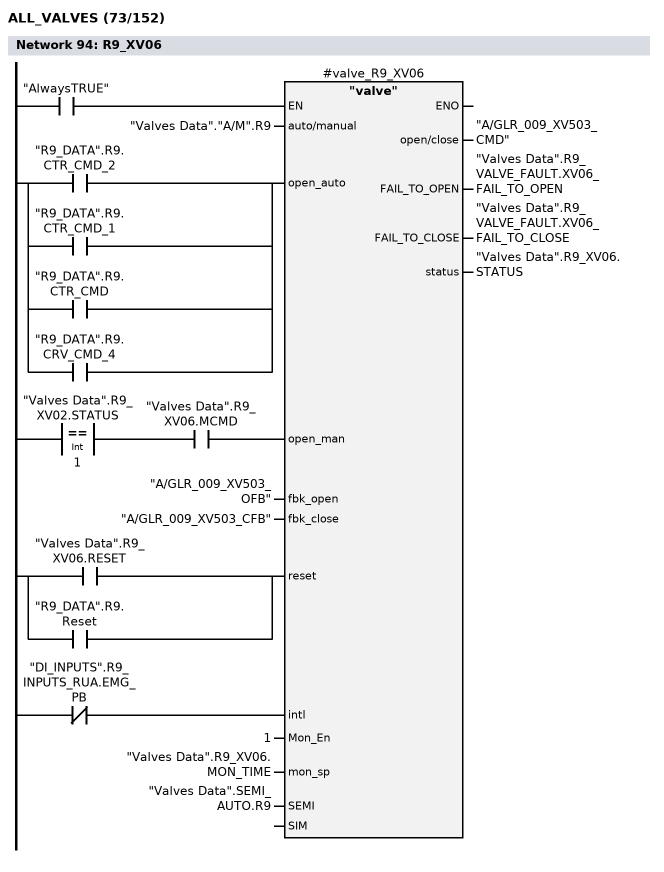
   RUNG wire#powerrail
      Contact( "AlwaysTRUE" )
      #valve_R9_XV06(open_auto := wire#w1, open_man := wire#w2, reset := wire#w3, intl := wire#w4, "auto/manual" := "Valves Data"."A/M".R9, fbk_open := "A/GLR_009_XV503_OFB", fbk_close := "A/GLR_009_XV503_CFB", Mon_En := 1, mon_sp := "Valves Data".R9_XV06.MON_TIME, SEMI := "Valves Data".SEMI_AUTO.R9, SIM :=, "open/close" => "A/GLR_009_XV503_CMD", FAIL_TO_OPEN => "Valves Data".R9_VALVE_FAULT.XV06_FAIL_TO_OPEN, FAIL_TO_CLOSE => "Valves Data".R9_VALVE_FAULT.XV06_FAIL_TO_CLOSE, status => "Valves Data".R9_XV06.STATUS)
   END_RUNG
   RUNG wire#powerrail
      Contact( "R9_DATA".R9.CTR_CMD_2 )
   END_RUNG wire#w1
   RUNG wire#powerrail
      Contact( "R9_DATA".R9.CTR_CMD_1 )
   END_RUNG wire#w1
   RUNG wire#powerrail
      Contact( "R9_DATA".R9.CTR_CMD )
   END_RUNG wire#w1
   RUNG wire#powerrail
      Contact( "R9_DATA".R9.CRV_CMD_4 )
   END_RUNG wire#w1
   RUNG wire#powerrail
      { S7_Templates := "SrcType := Int" } EQ_Contact(in1 := "Valves Data".R9_XV02.STATUS, in2 := 1)
      Contact( "Valves Data".R9_XV06.MCMD )
   END_RUNG wire#w2
   RUNG wire#powerrail
      Contact( "Valves Data".R9_XV06.RESET )
   END_RUNG wire#w3
   RUNG wire#powerrail
      Contact( "R9_DATA".R9.Reset )
   END_RUNG wire#w3
   RUNG wire#powerrail
      I_Contact( "DI_INPUTS".R9_INPUTS_RUA.EMG_PB )
   END_RUNG wire#w4
   // the same network as SCL:
   IF "AlwaysTRUE" THEN
       #valve_R9_XV06("auto/manual" := "Valves Data"."A/M".R9,   // "valve"
                      open_auto := "R9_DATA".R9.CTR_CMD_2 OR "R9_DATA".R9.CTR_CMD_1 OR "R9_DATA".R9.CTR_CMD OR "R9_DATA".R9.CRV_CMD_4,
                      open_man := ("Valves Data".R9_XV02.STATUS = 1) AND "Valves Data".R9_XV06.MCMD,
                      fbk_open := "A/GLR_009_XV503_OFB",
                      fbk_close := "A/GLR_009_XV503_CFB",
                      reset := "Valves Data".R9_XV06.RESET OR "R9_DATA".R9.Reset,
                      intl := NOT "DI_INPUTS".R9_INPUTS_RUA.EMG_PB,
                      Mon_En := 1,
                      mon_sp := "Valves Data".R9_XV06.MON_TIME,
                      SEMI := "Valves Data".SEMI_AUTO.R9,
                      "open/close" => "A/GLR_009_XV503_CMD",
                      FAIL_TO_OPEN => "Valves Data".R9_VALVE_FAULT.XV06_FAIL_TO_OPEN,
                      FAIL_TO_CLOSE => "Valves Data".R9_VALVE_FAULT.XV06_FAIL_TO_CLOSE,
                      status => "Valves Data".R9_XV06.STATUS);
   END_IF;
END_REGION

REGION Network 95: R9_XV07
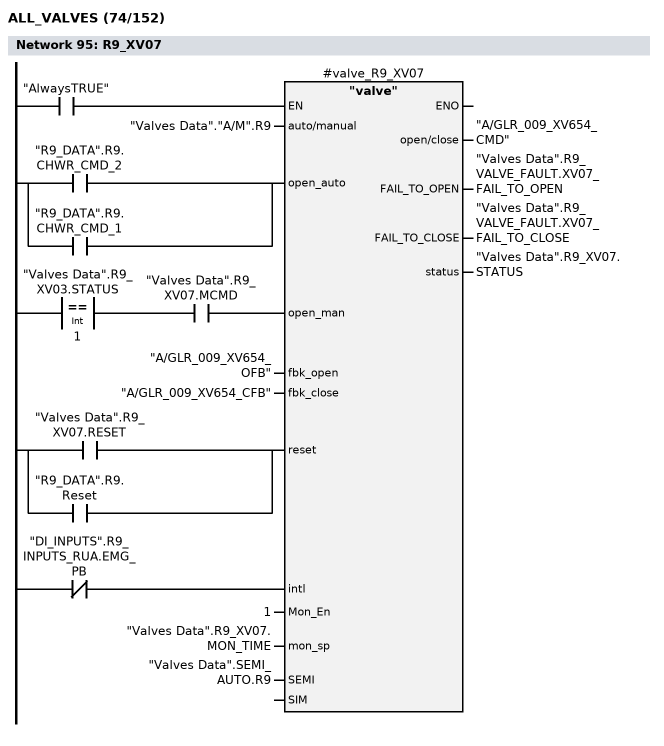
   RUNG wire#powerrail
      Contact( "AlwaysTRUE" )
      #valve_R9_XV07(open_auto := wire#w1, open_man := wire#w2, reset := wire#w3, intl := wire#w4, "auto/manual" := "Valves Data"."A/M".R9, fbk_open := "A/GLR_009_XV654_OFB", fbk_close := "A/GLR_009_XV654_CFB", Mon_En := 1, mon_sp := "Valves Data".R9_XV07.MON_TIME, SEMI := "Valves Data".SEMI_AUTO.R9, SIM :=, "open/close" => "A/GLR_009_XV654_CMD", FAIL_TO_OPEN => "Valves Data".R9_VALVE_FAULT.XV07_FAIL_TO_OPEN, FAIL_TO_CLOSE => "Valves Data".R9_VALVE_FAULT.XV07_FAIL_TO_CLOSE, status => "Valves Data".R9_XV07.STATUS)
   END_RUNG
   RUNG wire#powerrail
      Contact( "R9_DATA".R9.CHWR_CMD_2 )
   END_RUNG wire#w1
   RUNG wire#powerrail
      Contact( "R9_DATA".R9.CHWR_CMD_1 )
   END_RUNG wire#w1
   RUNG wire#powerrail
      { S7_Templates := "SrcType := Int" } EQ_Contact(in1 := "Valves Data".R9_XV03.STATUS, in2 := 1)
      Contact( "Valves Data".R9_XV07.MCMD )
   END_RUNG wire#w2
   RUNG wire#powerrail
      Contact( "Valves Data".R9_XV07.RESET )
   END_RUNG wire#w3
   RUNG wire#powerrail
      Contact( "R9_DATA".R9.Reset )
   END_RUNG wire#w3
   RUNG wire#powerrail
      I_Contact( "DI_INPUTS".R9_INPUTS_RUA.EMG_PB )
   END_RUNG wire#w4
   // the same network as SCL:
   IF "AlwaysTRUE" THEN
       #valve_R9_XV07("auto/manual" := "Valves Data"."A/M".R9,   // "valve"
                      open_auto := "R9_DATA".R9.CHWR_CMD_2 OR "R9_DATA".R9.CHWR_CMD_1,
                      open_man := ("Valves Data".R9_XV03.STATUS = 1) AND "Valves Data".R9_XV07.MCMD,
                      fbk_open := "A/GLR_009_XV654_OFB",
                      fbk_close := "A/GLR_009_XV654_CFB",
                      reset := "Valves Data".R9_XV07.RESET OR "R9_DATA".R9.Reset,
                      intl := NOT "DI_INPUTS".R9_INPUTS_RUA.EMG_PB,
                      Mon_En := 1,
                      mon_sp := "Valves Data".R9_XV07.MON_TIME,
                      SEMI := "Valves Data".SEMI_AUTO.R9,
                      "open/close" => "A/GLR_009_XV654_CMD",
                      FAIL_TO_OPEN => "Valves Data".R9_VALVE_FAULT.XV07_FAIL_TO_OPEN,
                      FAIL_TO_CLOSE => "Valves Data".R9_VALVE_FAULT.XV07_FAIL_TO_CLOSE,
                      status => "Valves Data".R9_XV07.STATUS);
   END_IF;
END_REGION

REGION Network 96: R9_XV08
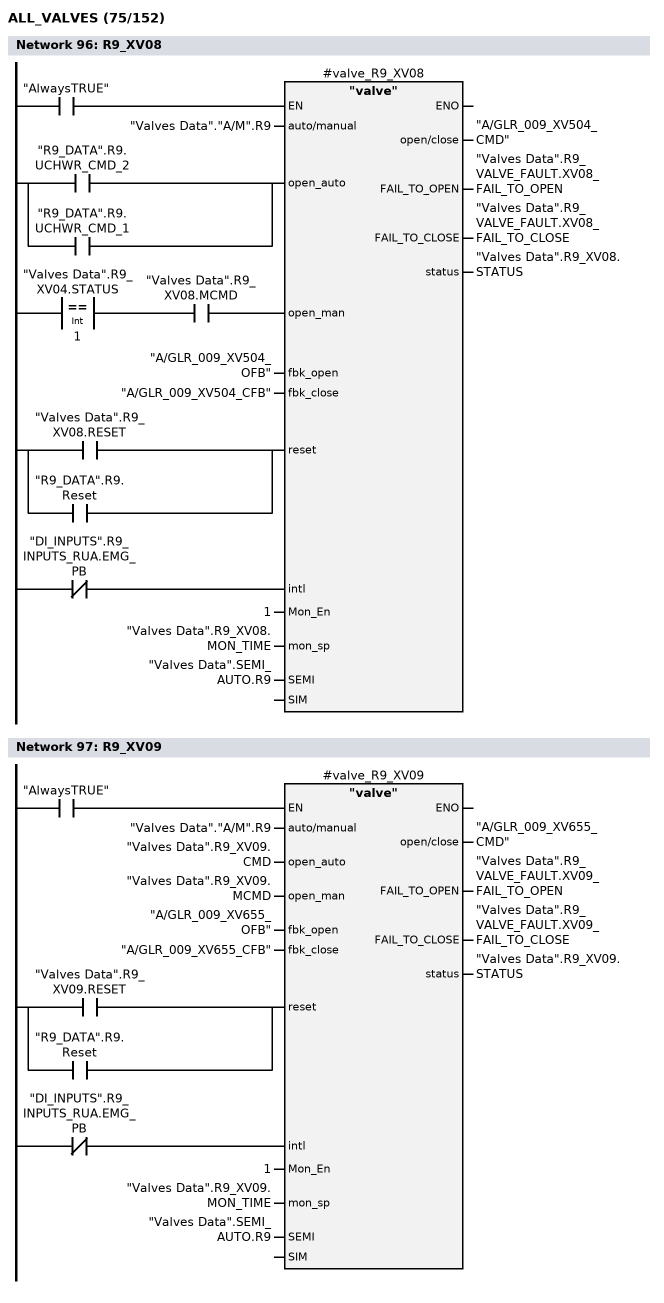
   RUNG wire#powerrail
      Contact( "AlwaysTRUE" )
      #valve_R9_XV08(open_auto := wire#w1, open_man := wire#w2, reset := wire#w3, intl := wire#w4, "auto/manual" := "Valves Data"."A/M".R9, fbk_open := "A/GLR_009_XV504_OFB", fbk_close := "A/GLR_009_XV504_CFB", Mon_En := 1, mon_sp := "Valves Data".R9_XV08.MON_TIME, SEMI := "Valves Data".SEMI_AUTO.R9, SIM :=, "open/close" => "A/GLR_009_XV504_CMD", FAIL_TO_OPEN => "Valves Data".R9_VALVE_FAULT.XV08_FAIL_TO_OPEN, FAIL_TO_CLOSE => "Valves Data".R9_VALVE_FAULT.XV08_FAIL_TO_CLOSE, status => "Valves Data".R9_XV08.STATUS)
   END_RUNG
   RUNG wire#powerrail
      Contact( "R9_DATA".R9.UCHWR_CMD_2 )
   END_RUNG wire#w1
   RUNG wire#powerrail
      Contact( "R9_DATA".R9.UCHWR_CMD_1 )
   END_RUNG wire#w1
   RUNG wire#powerrail
      { S7_Templates := "SrcType := Int" } EQ_Contact(in1 := "Valves Data".R9_XV04.STATUS, in2 := 1)
      Contact( "Valves Data".R9_XV08.MCMD )
   END_RUNG wire#w2
   RUNG wire#powerrail
      Contact( "Valves Data".R9_XV08.RESET )
   END_RUNG wire#w3
   RUNG wire#powerrail
      Contact( "R9_DATA".R9.Reset )
   END_RUNG wire#w3
   RUNG wire#powerrail
      I_Contact( "DI_INPUTS".R9_INPUTS_RUA.EMG_PB )
   END_RUNG wire#w4
   // the same network as SCL:
   IF "AlwaysTRUE" THEN
       #valve_R9_XV08("auto/manual" := "Valves Data"."A/M".R9,   // "valve"
                      open_auto := "R9_DATA".R9.UCHWR_CMD_2 OR "R9_DATA".R9.UCHWR_CMD_1,
                      open_man := ("Valves Data".R9_XV04.STATUS = 1) AND "Valves Data".R9_XV08.MCMD,
                      fbk_open := "A/GLR_009_XV504_OFB",
                      fbk_close := "A/GLR_009_XV504_CFB",
                      reset := "Valves Data".R9_XV08.RESET OR "R9_DATA".R9.Reset,
                      intl := NOT "DI_INPUTS".R9_INPUTS_RUA.EMG_PB,
                      Mon_En := 1,
                      mon_sp := "Valves Data".R9_XV08.MON_TIME,
                      SEMI := "Valves Data".SEMI_AUTO.R9,
                      "open/close" => "A/GLR_009_XV504_CMD",
                      FAIL_TO_OPEN => "Valves Data".R9_VALVE_FAULT.XV08_FAIL_TO_OPEN,
                      FAIL_TO_CLOSE => "Valves Data".R9_VALVE_FAULT.XV08_FAIL_TO_CLOSE,
                      status => "Valves Data".R9_XV08.STATUS);
   END_IF;
END_REGION

REGION Network 97: R9_XV09
   RUNG wire#powerrail
      Contact( "AlwaysTRUE" )
      #valve_R9_XV09(reset := wire#w1, intl := wire#w2, "auto/manual" := "Valves Data"."A/M".R9, open_auto := "Valves Data".R9_XV09.CMD, open_man := "Valves Data".R9_XV09.MCMD, fbk_open := "A/GLR_009_XV655_OFB", fbk_close := "A/GLR_009_XV655_CFB", Mon_En := 1, mon_sp := "Valves Data".R9_XV09.MON_TIME, SEMI := "Valves Data".SEMI_AUTO.R9, SIM :=, "open/close" => "A/GLR_009_XV655_CMD", FAIL_TO_OPEN => "Valves Data".R9_VALVE_FAULT.XV09_FAIL_TO_OPEN, FAIL_TO_CLOSE => "Valves Data".R9_VALVE_FAULT.XV09_FAIL_TO_CLOSE, status => "Valves Data".R9_XV09.STATUS)
   END_RUNG
   RUNG wire#powerrail
      Contact( "Valves Data".R9_XV09.RESET )
   END_RUNG wire#w1
   RUNG wire#powerrail
      Contact( "R9_DATA".R9.Reset )
   END_RUNG wire#w1
   RUNG wire#powerrail
      I_Contact( "DI_INPUTS".R9_INPUTS_RUA.EMG_PB )
   END_RUNG wire#w2
   // the same network as SCL:
   IF "AlwaysTRUE" THEN
       #valve_R9_XV09("auto/manual" := "Valves Data"."A/M".R9,   // "valve"
                      open_auto := "Valves Data".R9_XV09.CMD,
                      open_man := "Valves Data".R9_XV09.MCMD,
                      fbk_open := "A/GLR_009_XV655_OFB",
                      fbk_close := "A/GLR_009_XV655_CFB",
                      reset := "Valves Data".R9_XV09.RESET OR "R9_DATA".R9.Reset,
                      intl := NOT "DI_INPUTS".R9_INPUTS_RUA.EMG_PB,
                      Mon_En := 1,
                      mon_sp := "Valves Data".R9_XV09.MON_TIME,
                      SEMI := "Valves Data".SEMI_AUTO.R9,
                      "open/close" => "A/GLR_009_XV655_CMD",
                      FAIL_TO_OPEN => "Valves Data".R9_VALVE_FAULT.XV09_FAIL_TO_OPEN,
                      FAIL_TO_CLOSE => "Valves Data".R9_VALVE_FAULT.XV09_FAIL_TO_CLOSE,
                      status => "Valves Data".R9_XV09.STATUS);
   END_IF;
END_REGION

REGION Network 98: R9_XV10
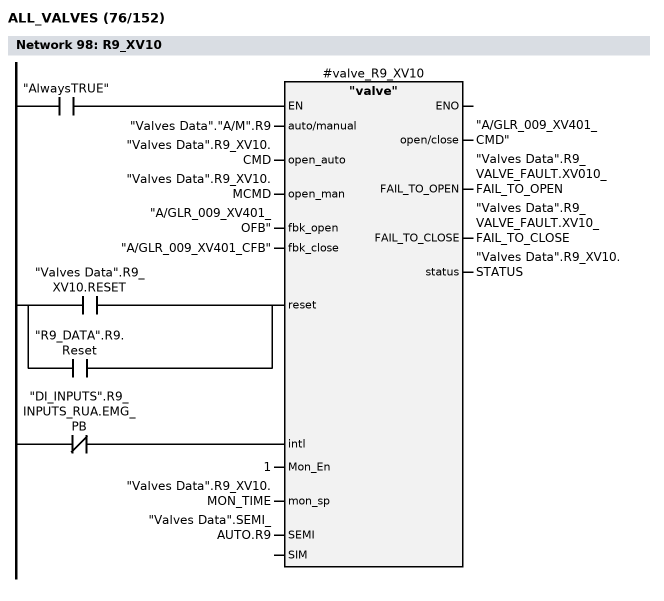
   RUNG wire#powerrail
      Contact( "AlwaysTRUE" )
      #valve_R9_XV10(reset := wire#w1, intl := wire#w2, "auto/manual" := "Valves Data"."A/M".R9, open_auto := "Valves Data".R9_XV10.CMD, open_man := "Valves Data".R9_XV10.MCMD, fbk_open := "A/GLR_009_XV401_OFB", fbk_close := "A/GLR_009_XV401_CFB", Mon_En := 1, mon_sp := "Valves Data".R9_XV10.MON_TIME, SEMI := "Valves Data".SEMI_AUTO.R9, SIM :=, "open/close" => "A/GLR_009_XV401_CMD", FAIL_TO_OPEN => "Valves Data".R9_VALVE_FAULT.XV010_FAIL_TO_OPEN, FAIL_TO_CLOSE => "Valves Data".R9_VALVE_FAULT.XV10_FAIL_TO_CLOSE, status => "Valves Data".R9_XV10.STATUS)
   END_RUNG
   RUNG wire#powerrail
      Contact( "Valves Data".R9_XV10.RESET )
   END_RUNG wire#w1
   RUNG wire#powerrail
      Contact( "R9_DATA".R9.Reset )
   END_RUNG wire#w1
   RUNG wire#powerrail
      I_Contact( "DI_INPUTS".R9_INPUTS_RUA.EMG_PB )
   END_RUNG wire#w2
   // the same network as SCL:
   IF "AlwaysTRUE" THEN
       #valve_R9_XV10("auto/manual" := "Valves Data"."A/M".R9,   // "valve"
                      open_auto := "Valves Data".R9_XV10.CMD,
                      open_man := "Valves Data".R9_XV10.MCMD,
                      fbk_open := "A/GLR_009_XV401_OFB",
                      fbk_close := "A/GLR_009_XV401_CFB",
                      reset := "Valves Data".R9_XV10.RESET OR "R9_DATA".R9.Reset,
                      intl := NOT "DI_INPUTS".R9_INPUTS_RUA.EMG_PB,
                      Mon_En := 1,
                      mon_sp := "Valves Data".R9_XV10.MON_TIME,
                      SEMI := "Valves Data".SEMI_AUTO.R9,
                      "open/close" => "A/GLR_009_XV401_CMD",
                      FAIL_TO_OPEN => "Valves Data".R9_VALVE_FAULT.XV010_FAIL_TO_OPEN,
                      FAIL_TO_CLOSE => "Valves Data".R9_VALVE_FAULT.XV10_FAIL_TO_CLOSE,
                      status => "Valves Data".R9_XV10.STATUS);
   END_IF;
END_REGION

REGION Network 99: ****REACTOR_10****
END_REGION

REGION Network 100: R10_XV01
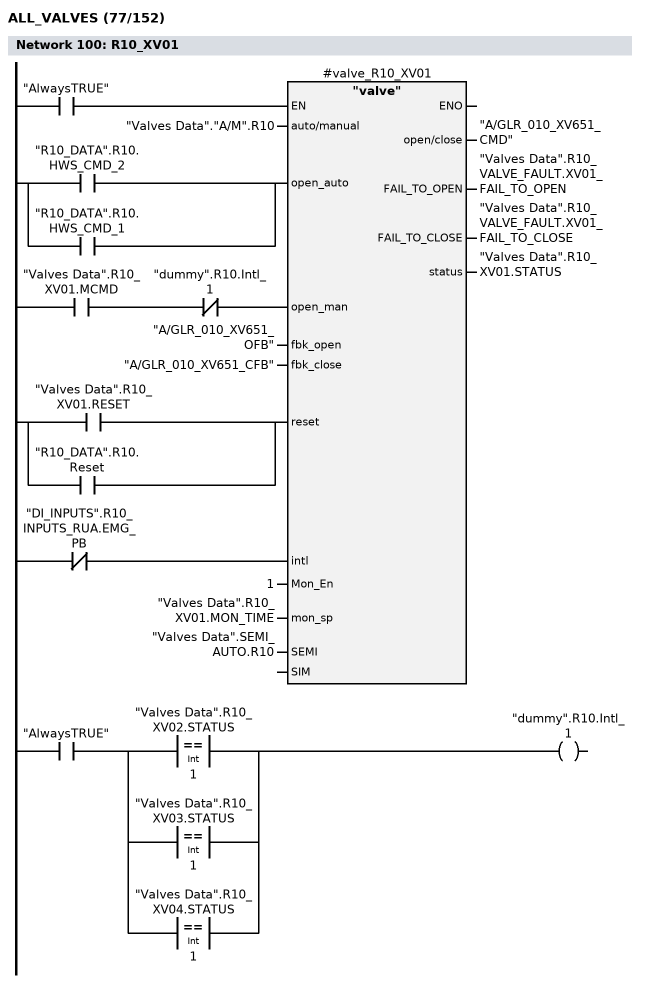
   RUNG wire#powerrail
      Contact( "AlwaysTRUE" )
      #valve_R10_XV01(open_auto := wire#w1, open_man := wire#w2, reset := wire#w3, intl := wire#w4, "auto/manual" := "Valves Data"."A/M".R10, fbk_open := "A/GLR_010_XV651_OFB", fbk_close := "A/GLR_010_XV651_CFB", Mon_En := 1, mon_sp := "Valves Data".R10_XV01.MON_TIME, SEMI := "Valves Data".SEMI_AUTO.R10, SIM :=, "open/close" => "A/GLR_010_XV651_CMD", FAIL_TO_OPEN => "Valves Data".R10_VALVE_FAULT.XV01_FAIL_TO_OPEN, FAIL_TO_CLOSE => "Valves Data".R10_VALVE_FAULT.XV01_FAIL_TO_CLOSE, status => "Valves Data".R10_XV01.STATUS)
   END_RUNG
   RUNG wire#powerrail
      Contact( "R10_DATA".R10.HWS_CMD_2 )
   END_RUNG wire#w1
   RUNG wire#powerrail
      Contact( "R10_DATA".R10.HWS_CMD_1 )
   END_RUNG wire#w1
   RUNG wire#powerrail
      Contact( "Valves Data".R10_XV01.MCMD )
      I_Contact( "dummy".R10.Intl_1 )
   END_RUNG wire#w2
   RUNG wire#powerrail
      Contact( "Valves Data".R10_XV01.RESET )
   END_RUNG wire#w3
   RUNG wire#powerrail
      Contact( "R10_DATA".R10.Reset )
   END_RUNG wire#w3
   RUNG wire#powerrail
      I_Contact( "DI_INPUTS".R10_INPUTS_RUA.EMG_PB )
   END_RUNG wire#w4
   RUNG wire#powerrail
      Contact( "AlwaysTRUE" )
      wire#w5
      { S7_Templates := "SrcType := Int" } EQ_Contact(in1 := "Valves Data".R10_XV02.STATUS, in2 := 1)
      wire#w6
      Coil( "dummy".R10.Intl_1 )
   END_RUNG
   RUNG wire#w5
      { S7_Templates := "SrcType := Int" } EQ_Contact(in1 := "Valves Data".R10_XV03.STATUS, in2 := 1)
   END_RUNG wire#w6
   RUNG wire#w5
      { S7_Templates := "SrcType := Int" } EQ_Contact(in1 := "Valves Data".R10_XV04.STATUS, in2 := 1)
   END_RUNG wire#w6
   // the same network as SCL:
   IF "AlwaysTRUE" THEN
       #valve_R10_XV01("auto/manual" := "Valves Data"."A/M".R10,   // "valve"
                       open_auto := "R10_DATA".R10.HWS_CMD_2 OR "R10_DATA".R10.HWS_CMD_1,
                       open_man := "Valves Data".R10_XV01.MCMD AND NOT "dummy".R10.Intl_1,
                       fbk_open := "A/GLR_010_XV651_OFB",
                       fbk_close := "A/GLR_010_XV651_CFB",
                       reset := "Valves Data".R10_XV01.RESET OR "R10_DATA".R10.Reset,
                       intl := NOT "DI_INPUTS".R10_INPUTS_RUA.EMG_PB,
                       Mon_En := 1,
                       mon_sp := "Valves Data".R10_XV01.MON_TIME,
                       SEMI := "Valves Data".SEMI_AUTO.R10,
                       "open/close" => "A/GLR_010_XV651_CMD",
                       FAIL_TO_OPEN => "Valves Data".R10_VALVE_FAULT.XV01_FAIL_TO_OPEN,
                       FAIL_TO_CLOSE => "Valves Data".R10_VALVE_FAULT.XV01_FAIL_TO_CLOSE,
                       status => "Valves Data".R10_XV01.STATUS);
   END_IF;
   "dummy".R10.Intl_1 := "AlwaysTRUE" AND (("Valves Data".R10_XV02.STATUS = 1) OR ("Valves Data".R10_XV03.STATUS = 1) OR ("Valves Data".R10_XV04.STATUS = 1));
END_REGION

REGION Network 101: R10_XV02
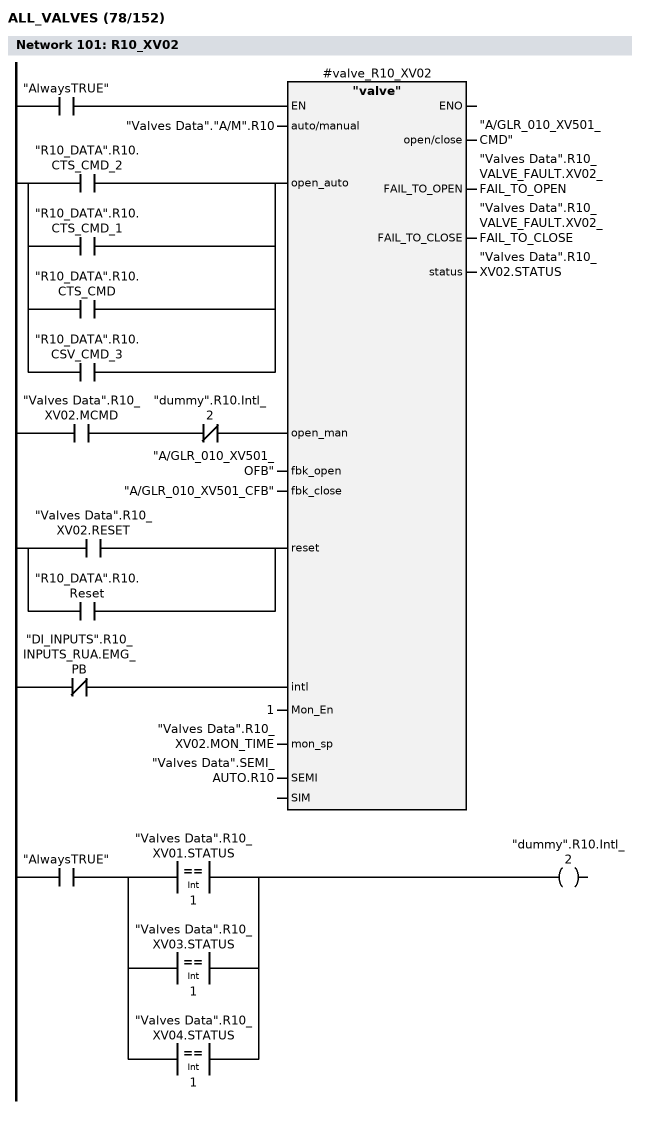
   RUNG wire#powerrail
      Contact( "AlwaysTRUE" )
      #valve_R10_XV02(open_auto := wire#w1, open_man := wire#w2, reset := wire#w3, intl := wire#w4, "auto/manual" := "Valves Data"."A/M".R10, fbk_open := "A/GLR_010_XV501_OFB", fbk_close := "A/GLR_010_XV501_CFB", Mon_En := 1, mon_sp := "Valves Data".R10_XV02.MON_TIME, SEMI := "Valves Data".SEMI_AUTO.R10, SIM :=, "open/close" => "A/GLR_010_XV501_CMD", FAIL_TO_OPEN => "Valves Data".R10_VALVE_FAULT.XV02_FAIL_TO_OPEN, FAIL_TO_CLOSE => "Valves Data".R10_VALVE_FAULT.XV02_FAIL_TO_CLOSE, status => "Valves Data".R10_XV02.STATUS)
   END_RUNG
   RUNG wire#powerrail
      Contact( "R10_DATA".R10.CTS_CMD_2 )
   END_RUNG wire#w1
   RUNG wire#powerrail
      Contact( "R10_DATA".R10.CTS_CMD_1 )
   END_RUNG wire#w1
   RUNG wire#powerrail
      Contact( "R10_DATA".R10.CTS_CMD )
   END_RUNG wire#w1
   RUNG wire#powerrail
      Contact( "R10_DATA".R10.CSV_CMD_3 )
   END_RUNG wire#w1
   RUNG wire#powerrail
      Contact( "Valves Data".R10_XV02.MCMD )
      I_Contact( "dummy".R10.Intl_2 )
   END_RUNG wire#w2
   RUNG wire#powerrail
      Contact( "Valves Data".R10_XV02.RESET )
   END_RUNG wire#w3
   RUNG wire#powerrail
      Contact( "R10_DATA".R10.Reset )
   END_RUNG wire#w3
   RUNG wire#powerrail
      I_Contact( "DI_INPUTS".R10_INPUTS_RUA.EMG_PB )
   END_RUNG wire#w4
   RUNG wire#powerrail
      Contact( "AlwaysTRUE" )
      wire#w5
      { S7_Templates := "SrcType := Int" } EQ_Contact(in1 := "Valves Data".R10_XV01.STATUS, in2 := 1)
      wire#w6
      Coil( "dummy".R10.Intl_2 )
   END_RUNG
   RUNG wire#w5
      { S7_Templates := "SrcType := Int" } EQ_Contact(in1 := "Valves Data".R10_XV03.STATUS, in2 := 1)
   END_RUNG wire#w6
   RUNG wire#w5
      { S7_Templates := "SrcType := Int" } EQ_Contact(in1 := "Valves Data".R10_XV04.STATUS, in2 := 1)
   END_RUNG wire#w6
   // the same network as SCL:
   IF "AlwaysTRUE" THEN
       #valve_R10_XV02("auto/manual" := "Valves Data"."A/M".R10,   // "valve"
                       open_auto := "R10_DATA".R10.CTS_CMD_2 OR "R10_DATA".R10.CTS_CMD_1 OR "R10_DATA".R10.CTS_CMD OR "R10_DATA".R10.CSV_CMD_3,
                       open_man := "Valves Data".R10_XV02.MCMD AND NOT "dummy".R10.Intl_2,
                       fbk_open := "A/GLR_010_XV501_OFB",
                       fbk_close := "A/GLR_010_XV501_CFB",
                       reset := "Valves Data".R10_XV02.RESET OR "R10_DATA".R10.Reset,
                       intl := NOT "DI_INPUTS".R10_INPUTS_RUA.EMG_PB,
                       Mon_En := 1,
                       mon_sp := "Valves Data".R10_XV02.MON_TIME,
                       SEMI := "Valves Data".SEMI_AUTO.R10,
                       "open/close" => "A/GLR_010_XV501_CMD",
                       FAIL_TO_OPEN => "Valves Data".R10_VALVE_FAULT.XV02_FAIL_TO_OPEN,
                       FAIL_TO_CLOSE => "Valves Data".R10_VALVE_FAULT.XV02_FAIL_TO_CLOSE,
                       status => "Valves Data".R10_XV02.STATUS);
   END_IF;
   "dummy".R10.Intl_2 := "AlwaysTRUE" AND (("Valves Data".R10_XV01.STATUS = 1) OR ("Valves Data".R10_XV03.STATUS = 1) OR ("Valves Data".R10_XV04.STATUS = 1));
END_REGION

REGION Network 102: R10_XV03
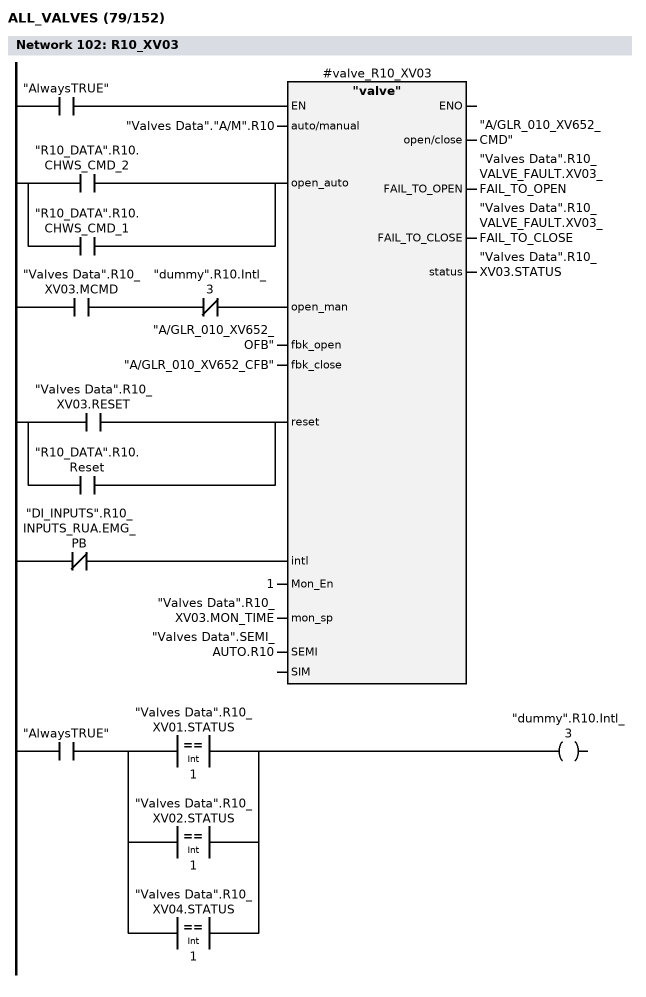
   RUNG wire#powerrail
      Contact( "AlwaysTRUE" )
      #valve_R10_XV03(open_auto := wire#w1, open_man := wire#w2, reset := wire#w3, intl := wire#w4, "auto/manual" := "Valves Data"."A/M".R10, fbk_open := "A/GLR_010_XV652_OFB", fbk_close := "A/GLR_010_XV652_CFB", Mon_En := 1, mon_sp := "Valves Data".R10_XV03.MON_TIME, SEMI := "Valves Data".SEMI_AUTO.R10, SIM :=, "open/close" => "A/GLR_010_XV652_CMD", FAIL_TO_OPEN => "Valves Data".R10_VALVE_FAULT.XV03_FAIL_TO_OPEN, FAIL_TO_CLOSE => "Valves Data".R10_VALVE_FAULT.XV03_FAIL_TO_CLOSE, status => "Valves Data".R10_XV03.STATUS)
   END_RUNG
   RUNG wire#powerrail
      Contact( "R10_DATA".R10.CHWS_CMD_2 )
   END_RUNG wire#w1
   RUNG wire#powerrail
      Contact( "R10_DATA".R10.CHWS_CMD_1 )
   END_RUNG wire#w1
   RUNG wire#powerrail
      Contact( "Valves Data".R10_XV03.MCMD )
      I_Contact( "dummy".R10.Intl_3 )
   END_RUNG wire#w2
   RUNG wire#powerrail
      Contact( "Valves Data".R10_XV03.RESET )
   END_RUNG wire#w3
   RUNG wire#powerrail
      Contact( "R10_DATA".R10.Reset )
   END_RUNG wire#w3
   RUNG wire#powerrail
      I_Contact( "DI_INPUTS".R10_INPUTS_RUA.EMG_PB )
   END_RUNG wire#w4
   RUNG wire#powerrail
      Contact( "AlwaysTRUE" )
      wire#w5
      { S7_Templates := "SrcType := Int" } EQ_Contact(in1 := "Valves Data".R10_XV01.STATUS, in2 := 1)
      wire#w6
      Coil( "dummy".R10.Intl_3 )
   END_RUNG
   RUNG wire#w5
      { S7_Templates := "SrcType := Int" } EQ_Contact(in1 := "Valves Data".R10_XV02.STATUS, in2 := 1)
   END_RUNG wire#w6
   RUNG wire#w5
      { S7_Templates := "SrcType := Int" } EQ_Contact(in1 := "Valves Data".R10_XV04.STATUS, in2 := 1)
   END_RUNG wire#w6
   // the same network as SCL:
   IF "AlwaysTRUE" THEN
       #valve_R10_XV03("auto/manual" := "Valves Data"."A/M".R10,   // "valve"
                       open_auto := "R10_DATA".R10.CHWS_CMD_2 OR "R10_DATA".R10.CHWS_CMD_1,
                       open_man := "Valves Data".R10_XV03.MCMD AND NOT "dummy".R10.Intl_3,
                       fbk_open := "A/GLR_010_XV652_OFB",
                       fbk_close := "A/GLR_010_XV652_CFB",
                       reset := "Valves Data".R10_XV03.RESET OR "R10_DATA".R10.Reset,
                       intl := NOT "DI_INPUTS".R10_INPUTS_RUA.EMG_PB,
                       Mon_En := 1,
                       mon_sp := "Valves Data".R10_XV03.MON_TIME,
                       SEMI := "Valves Data".SEMI_AUTO.R10,
                       "open/close" => "A/GLR_010_XV652_CMD",
                       FAIL_TO_OPEN => "Valves Data".R10_VALVE_FAULT.XV03_FAIL_TO_OPEN,
                       FAIL_TO_CLOSE => "Valves Data".R10_VALVE_FAULT.XV03_FAIL_TO_CLOSE,
                       status => "Valves Data".R10_XV03.STATUS);
   END_IF;
   "dummy".R10.Intl_3 := "AlwaysTRUE" AND (("Valves Data".R10_XV01.STATUS = 1) OR ("Valves Data".R10_XV02.STATUS = 1) OR ("Valves Data".R10_XV04.STATUS = 1));
END_REGION

REGION Network 103: R10_XV04
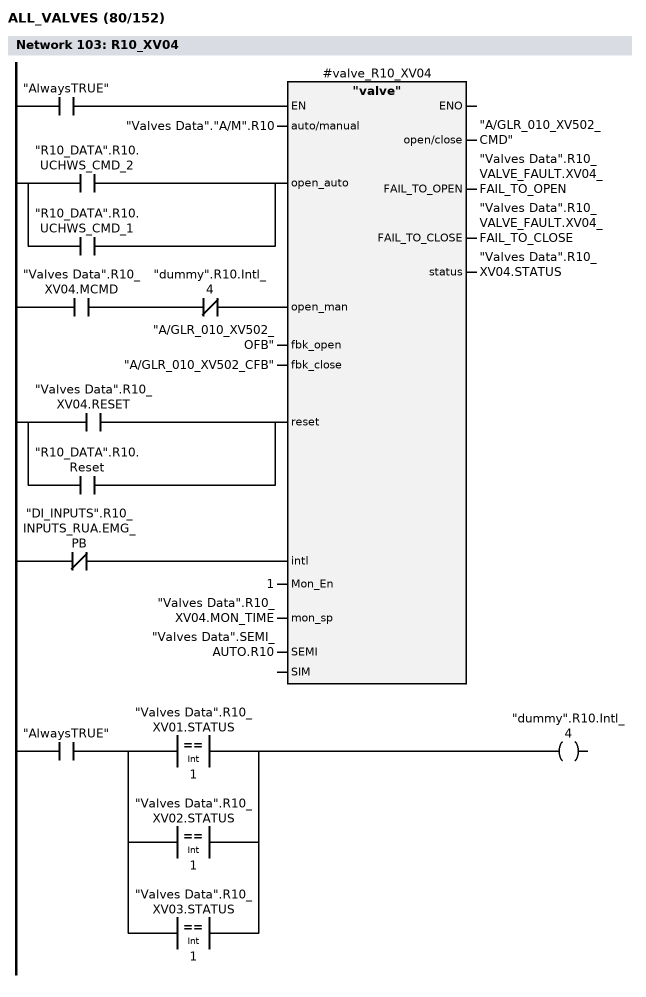
   RUNG wire#powerrail
      Contact( "AlwaysTRUE" )
      #valve_R10_XV04(open_auto := wire#w1, open_man := wire#w2, reset := wire#w3, intl := wire#w4, "auto/manual" := "Valves Data"."A/M".R10, fbk_open := "A/GLR_010_XV502_OFB", fbk_close := "A/GLR_010_XV502_CFB", Mon_En := 1, mon_sp := "Valves Data".R10_XV04.MON_TIME, SEMI := "Valves Data".SEMI_AUTO.R10, SIM :=, "open/close" => "A/GLR_010_XV502_CMD", FAIL_TO_OPEN => "Valves Data".R10_VALVE_FAULT.XV04_FAIL_TO_OPEN, FAIL_TO_CLOSE => "Valves Data".R10_VALVE_FAULT.XV04_FAIL_TO_CLOSE, status => "Valves Data".R10_XV04.STATUS)
   END_RUNG
   RUNG wire#powerrail
      Contact( "R10_DATA".R10.UCHWS_CMD_2 )
   END_RUNG wire#w1
   RUNG wire#powerrail
      Contact( "R10_DATA".R10.UCHWS_CMD_1 )
   END_RUNG wire#w1
   RUNG wire#powerrail
      Contact( "Valves Data".R10_XV04.MCMD )
      I_Contact( "dummy".R10.Intl_4 )
   END_RUNG wire#w2
   RUNG wire#powerrail
      Contact( "Valves Data".R10_XV04.RESET )
   END_RUNG wire#w3
   RUNG wire#powerrail
      Contact( "R10_DATA".R10.Reset )
   END_RUNG wire#w3
   RUNG wire#powerrail
      I_Contact( "DI_INPUTS".R10_INPUTS_RUA.EMG_PB )
   END_RUNG wire#w4
   RUNG wire#powerrail
      Contact( "AlwaysTRUE" )
      wire#w5
      { S7_Templates := "SrcType := Int" } EQ_Contact(in1 := "Valves Data".R10_XV01.STATUS, in2 := 1)
      wire#w6
      Coil( "dummy".R10.Intl_4 )
   END_RUNG
   RUNG wire#w5
      { S7_Templates := "SrcType := Int" } EQ_Contact(in1 := "Valves Data".R10_XV02.STATUS, in2 := 1)
   END_RUNG wire#w6
   RUNG wire#w5
      { S7_Templates := "SrcType := Int" } EQ_Contact(in1 := "Valves Data".R10_XV03.STATUS, in2 := 1)
   END_RUNG wire#w6
   // the same network as SCL:
   IF "AlwaysTRUE" THEN
       #valve_R10_XV04("auto/manual" := "Valves Data"."A/M".R10,   // "valve"
                       open_auto := "R10_DATA".R10.UCHWS_CMD_2 OR "R10_DATA".R10.UCHWS_CMD_1,
                       open_man := "Valves Data".R10_XV04.MCMD AND NOT "dummy".R10.Intl_4,
                       fbk_open := "A/GLR_010_XV502_OFB",
                       fbk_close := "A/GLR_010_XV502_CFB",
                       reset := "Valves Data".R10_XV04.RESET OR "R10_DATA".R10.Reset,
                       intl := NOT "DI_INPUTS".R10_INPUTS_RUA.EMG_PB,
                       Mon_En := 1,
                       mon_sp := "Valves Data".R10_XV04.MON_TIME,
                       SEMI := "Valves Data".SEMI_AUTO.R10,
                       "open/close" => "A/GLR_010_XV502_CMD",
                       FAIL_TO_OPEN => "Valves Data".R10_VALVE_FAULT.XV04_FAIL_TO_OPEN,
                       FAIL_TO_CLOSE => "Valves Data".R10_VALVE_FAULT.XV04_FAIL_TO_CLOSE,
                       status => "Valves Data".R10_XV04.STATUS);
   END_IF;
   "dummy".R10.Intl_4 := "AlwaysTRUE" AND (("Valves Data".R10_XV01.STATUS = 1) OR ("Valves Data".R10_XV02.STATUS = 1) OR ("Valves Data".R10_XV03.STATUS = 1));
END_REGION

REGION Network 104: R10_XV05
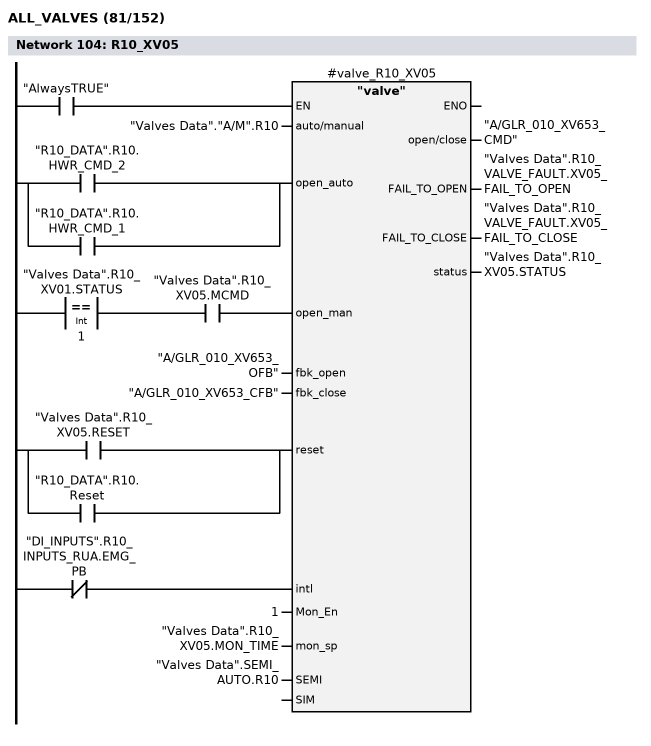
   RUNG wire#powerrail
      Contact( "AlwaysTRUE" )
      #valve_R10_XV05(open_auto := wire#w1, open_man := wire#w2, reset := wire#w3, intl := wire#w4, "auto/manual" := "Valves Data"."A/M".R10, fbk_open := "A/GLR_010_XV653_OFB", fbk_close := "A/GLR_010_XV653_CFB", Mon_En := 1, mon_sp := "Valves Data".R10_XV05.MON_TIME, SEMI := "Valves Data".SEMI_AUTO.R10, SIM :=, "open/close" => "A/GLR_010_XV653_CMD", FAIL_TO_OPEN => "Valves Data".R10_VALVE_FAULT.XV05_FAIL_TO_OPEN, FAIL_TO_CLOSE => "Valves Data".R10_VALVE_FAULT.XV05_FAIL_TO_CLOSE, status => "Valves Data".R10_XV05.STATUS)
   END_RUNG
   RUNG wire#powerrail
      Contact( "R10_DATA".R10.HWR_CMD_2 )
   END_RUNG wire#w1
   RUNG wire#powerrail
      Contact( "R10_DATA".R10.HWR_CMD_1 )
   END_RUNG wire#w1
   RUNG wire#powerrail
      { S7_Templates := "SrcType := Int" } EQ_Contact(in1 := "Valves Data".R10_XV01.STATUS, in2 := 1)
      Contact( "Valves Data".R10_XV05.MCMD )
   END_RUNG wire#w2
   RUNG wire#powerrail
      Contact( "Valves Data".R10_XV05.RESET )
   END_RUNG wire#w3
   RUNG wire#powerrail
      Contact( "R10_DATA".R10.Reset )
   END_RUNG wire#w3
   RUNG wire#powerrail
      I_Contact( "DI_INPUTS".R10_INPUTS_RUA.EMG_PB )
   END_RUNG wire#w4
   // the same network as SCL:
   IF "AlwaysTRUE" THEN
       #valve_R10_XV05("auto/manual" := "Valves Data"."A/M".R10,   // "valve"
                       open_auto := "R10_DATA".R10.HWR_CMD_2 OR "R10_DATA".R10.HWR_CMD_1,
                       open_man := ("Valves Data".R10_XV01.STATUS = 1) AND "Valves Data".R10_XV05.MCMD,
                       fbk_open := "A/GLR_010_XV653_OFB",
                       fbk_close := "A/GLR_010_XV653_CFB",
                       reset := "Valves Data".R10_XV05.RESET OR "R10_DATA".R10.Reset,
                       intl := NOT "DI_INPUTS".R10_INPUTS_RUA.EMG_PB,
                       Mon_En := 1,
                       mon_sp := "Valves Data".R10_XV05.MON_TIME,
                       SEMI := "Valves Data".SEMI_AUTO.R10,
                       "open/close" => "A/GLR_010_XV653_CMD",
                       FAIL_TO_OPEN => "Valves Data".R10_VALVE_FAULT.XV05_FAIL_TO_OPEN,
                       FAIL_TO_CLOSE => "Valves Data".R10_VALVE_FAULT.XV05_FAIL_TO_CLOSE,
                       status => "Valves Data".R10_XV05.STATUS);
   END_IF;
END_REGION

REGION Network 105: R10_XV06
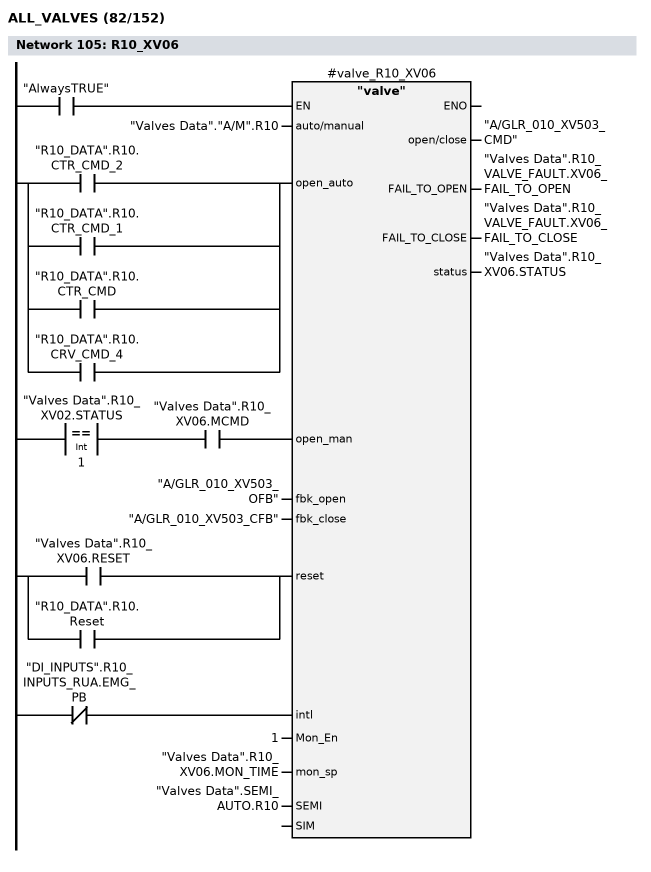
   RUNG wire#powerrail
      Contact( "AlwaysTRUE" )
      #valve_R10_XV06(open_auto := wire#w1, open_man := wire#w2, reset := wire#w3, intl := wire#w4, "auto/manual" := "Valves Data"."A/M".R10, fbk_open := "A/GLR_010_XV503_OFB", fbk_close := "A/GLR_010_XV503_CFB", Mon_En := 1, mon_sp := "Valves Data".R10_XV06.MON_TIME, SEMI := "Valves Data".SEMI_AUTO.R10, SIM :=, "open/close" => "A/GLR_010_XV503_CMD", FAIL_TO_OPEN => "Valves Data".R10_VALVE_FAULT.XV06_FAIL_TO_OPEN, FAIL_TO_CLOSE => "Valves Data".R10_VALVE_FAULT.XV06_FAIL_TO_CLOSE, status => "Valves Data".R10_XV06.STATUS)
   END_RUNG
   RUNG wire#powerrail
      Contact( "R10_DATA".R10.CTR_CMD_2 )
   END_RUNG wire#w1
   RUNG wire#powerrail
      Contact( "R10_DATA".R10.CTR_CMD_1 )
   END_RUNG wire#w1
   RUNG wire#powerrail
      Contact( "R10_DATA".R10.CTR_CMD )
   END_RUNG wire#w1
   RUNG wire#powerrail
      Contact( "R10_DATA".R10.CRV_CMD_4 )
   END_RUNG wire#w1
   RUNG wire#powerrail
      { S7_Templates := "SrcType := Int" } EQ_Contact(in1 := "Valves Data".R10_XV02.STATUS, in2 := 1)
      Contact( "Valves Data".R10_XV06.MCMD )
   END_RUNG wire#w2
   RUNG wire#powerrail
      Contact( "Valves Data".R10_XV06.RESET )
   END_RUNG wire#w3
   RUNG wire#powerrail
      Contact( "R10_DATA".R10.Reset )
   END_RUNG wire#w3
   RUNG wire#powerrail
      I_Contact( "DI_INPUTS".R10_INPUTS_RUA.EMG_PB )
   END_RUNG wire#w4
   // the same network as SCL:
   IF "AlwaysTRUE" THEN
       #valve_R10_XV06("auto/manual" := "Valves Data"."A/M".R10,   // "valve"
                       open_auto := "R10_DATA".R10.CTR_CMD_2 OR "R10_DATA".R10.CTR_CMD_1 OR "R10_DATA".R10.CTR_CMD OR "R10_DATA".R10.CRV_CMD_4,
                       open_man := ("Valves Data".R10_XV02.STATUS = 1) AND "Valves Data".R10_XV06.MCMD,
                       fbk_open := "A/GLR_010_XV503_OFB",
                       fbk_close := "A/GLR_010_XV503_CFB",
                       reset := "Valves Data".R10_XV06.RESET OR "R10_DATA".R10.Reset,
                       intl := NOT "DI_INPUTS".R10_INPUTS_RUA.EMG_PB,
                       Mon_En := 1,
                       mon_sp := "Valves Data".R10_XV06.MON_TIME,
                       SEMI := "Valves Data".SEMI_AUTO.R10,
                       "open/close" => "A/GLR_010_XV503_CMD",
                       FAIL_TO_OPEN => "Valves Data".R10_VALVE_FAULT.XV06_FAIL_TO_OPEN,
                       FAIL_TO_CLOSE => "Valves Data".R10_VALVE_FAULT.XV06_FAIL_TO_CLOSE,
                       status => "Valves Data".R10_XV06.STATUS);
   END_IF;
END_REGION

REGION Network 106: R10_XV07
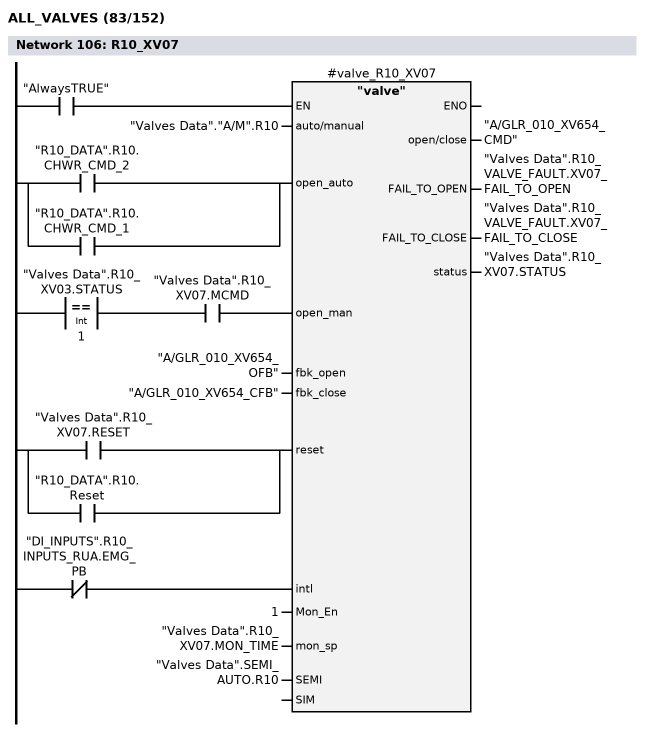
   RUNG wire#powerrail
      Contact( "AlwaysTRUE" )
      #valve_R10_XV07(open_auto := wire#w1, open_man := wire#w2, reset := wire#w3, intl := wire#w4, "auto/manual" := "Valves Data"."A/M".R10, fbk_open := "A/GLR_010_XV654_OFB", fbk_close := "A/GLR_010_XV654_CFB", Mon_En := 1, mon_sp := "Valves Data".R10_XV07.MON_TIME, SEMI := "Valves Data".SEMI_AUTO.R10, SIM :=, "open/close" => "A/GLR_010_XV654_CMD", FAIL_TO_OPEN => "Valves Data".R10_VALVE_FAULT.XV07_FAIL_TO_OPEN, FAIL_TO_CLOSE => "Valves Data".R10_VALVE_FAULT.XV07_FAIL_TO_CLOSE, status => "Valves Data".R10_XV07.STATUS)
   END_RUNG
   RUNG wire#powerrail
      Contact( "R10_DATA".R10.CHWR_CMD_2 )
   END_RUNG wire#w1
   RUNG wire#powerrail
      Contact( "R10_DATA".R10.CHWR_CMD_1 )
   END_RUNG wire#w1
   RUNG wire#powerrail
      { S7_Templates := "SrcType := Int" } EQ_Contact(in1 := "Valves Data".R10_XV03.STATUS, in2 := 1)
      Contact( "Valves Data".R10_XV07.MCMD )
   END_RUNG wire#w2
   RUNG wire#powerrail
      Contact( "Valves Data".R10_XV07.RESET )
   END_RUNG wire#w3
   RUNG wire#powerrail
      Contact( "R10_DATA".R10.Reset )
   END_RUNG wire#w3
   RUNG wire#powerrail
      I_Contact( "DI_INPUTS".R10_INPUTS_RUA.EMG_PB )
   END_RUNG wire#w4
   // the same network as SCL:
   IF "AlwaysTRUE" THEN
       #valve_R10_XV07("auto/manual" := "Valves Data"."A/M".R10,   // "valve"
                       open_auto := "R10_DATA".R10.CHWR_CMD_2 OR "R10_DATA".R10.CHWR_CMD_1,
                       open_man := ("Valves Data".R10_XV03.STATUS = 1) AND "Valves Data".R10_XV07.MCMD,
                       fbk_open := "A/GLR_010_XV654_OFB",
                       fbk_close := "A/GLR_010_XV654_CFB",
                       reset := "Valves Data".R10_XV07.RESET OR "R10_DATA".R10.Reset,
                       intl := NOT "DI_INPUTS".R10_INPUTS_RUA.EMG_PB,
                       Mon_En := 1,
                       mon_sp := "Valves Data".R10_XV07.MON_TIME,
                       SEMI := "Valves Data".SEMI_AUTO.R10,
                       "open/close" => "A/GLR_010_XV654_CMD",
                       FAIL_TO_OPEN => "Valves Data".R10_VALVE_FAULT.XV07_FAIL_TO_OPEN,
                       FAIL_TO_CLOSE => "Valves Data".R10_VALVE_FAULT.XV07_FAIL_TO_CLOSE,
                       status => "Valves Data".R10_XV07.STATUS);
   END_IF;
END_REGION

REGION Network 107: R10_XV08
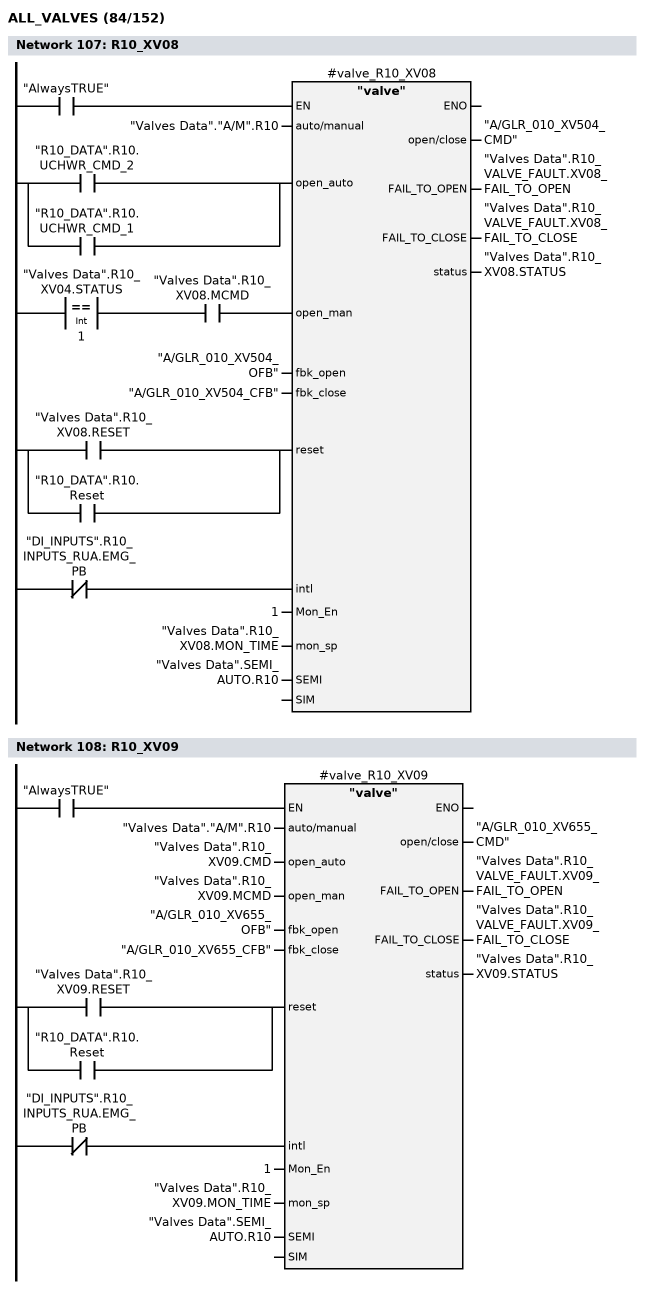
   RUNG wire#powerrail
      Contact( "AlwaysTRUE" )
      #valve_R10_XV08(open_auto := wire#w1, open_man := wire#w2, reset := wire#w3, intl := wire#w4, "auto/manual" := "Valves Data"."A/M".R10, fbk_open := "A/GLR_010_XV504_OFB", fbk_close := "A/GLR_010_XV504_CFB", Mon_En := 1, mon_sp := "Valves Data".R10_XV08.MON_TIME, SEMI := "Valves Data".SEMI_AUTO.R10, SIM :=, "open/close" => "A/GLR_010_XV504_CMD", FAIL_TO_OPEN => "Valves Data".R10_VALVE_FAULT.XV08_FAIL_TO_OPEN, FAIL_TO_CLOSE => "Valves Data".R10_VALVE_FAULT.XV08_FAIL_TO_CLOSE, status => "Valves Data".R10_XV08.STATUS)
   END_RUNG
   RUNG wire#powerrail
      Contact( "R10_DATA".R10.UCHWR_CMD_2 )
   END_RUNG wire#w1
   RUNG wire#powerrail
      Contact( "R10_DATA".R10.UCHWR_CMD_1 )
   END_RUNG wire#w1
   RUNG wire#powerrail
      { S7_Templates := "SrcType := Int" } EQ_Contact(in1 := "Valves Data".R10_XV04.STATUS, in2 := 1)
      Contact( "Valves Data".R10_XV08.MCMD )
   END_RUNG wire#w2
   RUNG wire#powerrail
      Contact( "Valves Data".R10_XV08.RESET )
   END_RUNG wire#w3
   RUNG wire#powerrail
      Contact( "R10_DATA".R10.Reset )
   END_RUNG wire#w3
   RUNG wire#powerrail
      I_Contact( "DI_INPUTS".R10_INPUTS_RUA.EMG_PB )
   END_RUNG wire#w4
   // the same network as SCL:
   IF "AlwaysTRUE" THEN
       #valve_R10_XV08("auto/manual" := "Valves Data"."A/M".R10,   // "valve"
                       open_auto := "R10_DATA".R10.UCHWR_CMD_2 OR "R10_DATA".R10.UCHWR_CMD_1,
                       open_man := ("Valves Data".R10_XV04.STATUS = 1) AND "Valves Data".R10_XV08.MCMD,
                       fbk_open := "A/GLR_010_XV504_OFB",
                       fbk_close := "A/GLR_010_XV504_CFB",
                       reset := "Valves Data".R10_XV08.RESET OR "R10_DATA".R10.Reset,
                       intl := NOT "DI_INPUTS".R10_INPUTS_RUA.EMG_PB,
                       Mon_En := 1,
                       mon_sp := "Valves Data".R10_XV08.MON_TIME,
                       SEMI := "Valves Data".SEMI_AUTO.R10,
                       "open/close" => "A/GLR_010_XV504_CMD",
                       FAIL_TO_OPEN => "Valves Data".R10_VALVE_FAULT.XV08_FAIL_TO_OPEN,
                       FAIL_TO_CLOSE => "Valves Data".R10_VALVE_FAULT.XV08_FAIL_TO_CLOSE,
                       status => "Valves Data".R10_XV08.STATUS);
   END_IF;
END_REGION

REGION Network 108: R10_XV09
   RUNG wire#powerrail
      Contact( "AlwaysTRUE" )
      #valve_R10_XV09(reset := wire#w1, intl := wire#w2, "auto/manual" := "Valves Data"."A/M".R10, open_auto := "Valves Data".R10_XV09.CMD, open_man := "Valves Data".R10_XV09.MCMD, fbk_open := "A/GLR_010_XV655_OFB", fbk_close := "A/GLR_010_XV655_CFB", Mon_En := 1, mon_sp := "Valves Data".R10_XV09.MON_TIME, SEMI := "Valves Data".SEMI_AUTO.R10, SIM :=, "open/close" => "A/GLR_010_XV655_CMD", FAIL_TO_OPEN => "Valves Data".R10_VALVE_FAULT.XV09_FAIL_TO_OPEN, FAIL_TO_CLOSE => "Valves Data".R10_VALVE_FAULT.XV09_FAIL_TO_CLOSE, status => "Valves Data".R10_XV09.STATUS)
   END_RUNG
   RUNG wire#powerrail
      Contact( "Valves Data".R10_XV09.RESET )
   END_RUNG wire#w1
   RUNG wire#powerrail
      Contact( "R10_DATA".R10.Reset )
   END_RUNG wire#w1
   RUNG wire#powerrail
      I_Contact( "DI_INPUTS".R10_INPUTS_RUA.EMG_PB )
   END_RUNG wire#w2
   // the same network as SCL:
   IF "AlwaysTRUE" THEN
       #valve_R10_XV09("auto/manual" := "Valves Data"."A/M".R10,   // "valve"
                       open_auto := "Valves Data".R10_XV09.CMD,
                       open_man := "Valves Data".R10_XV09.MCMD,
                       fbk_open := "A/GLR_010_XV655_OFB",
                       fbk_close := "A/GLR_010_XV655_CFB",
                       reset := "Valves Data".R10_XV09.RESET OR "R10_DATA".R10.Reset,
                       intl := NOT "DI_INPUTS".R10_INPUTS_RUA.EMG_PB,
                       Mon_En := 1,
                       mon_sp := "Valves Data".R10_XV09.MON_TIME,
                       SEMI := "Valves Data".SEMI_AUTO.R10,
                       "open/close" => "A/GLR_010_XV655_CMD",
                       FAIL_TO_OPEN => "Valves Data".R10_VALVE_FAULT.XV09_FAIL_TO_OPEN,
                       FAIL_TO_CLOSE => "Valves Data".R10_VALVE_FAULT.XV09_FAIL_TO_CLOSE,
                       status => "Valves Data".R10_XV09.STATUS);
   END_IF;
END_REGION

REGION Network 109: R10_XV10
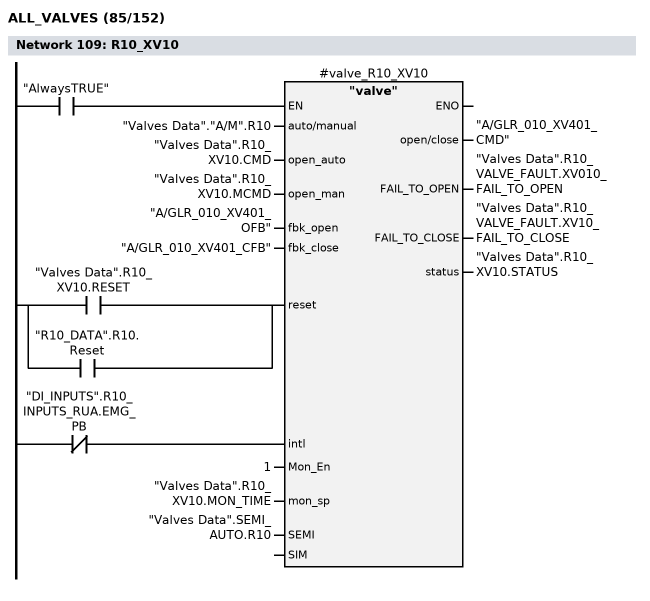
   RUNG wire#powerrail
      Contact( "AlwaysTRUE" )
      #valve_R10_XV10(reset := wire#w1, intl := wire#w2, "auto/manual" := "Valves Data"."A/M".R10, open_auto := "Valves Data".R10_XV10.CMD, open_man := "Valves Data".R10_XV10.MCMD, fbk_open := "A/GLR_010_XV401_OFB", fbk_close := "A/GLR_010_XV401_CFB", Mon_En := 1, mon_sp := "Valves Data".R10_XV10.MON_TIME, SEMI := "Valves Data".SEMI_AUTO.R10, SIM :=, "open/close" => "A/GLR_010_XV401_CMD", FAIL_TO_OPEN => "Valves Data".R10_VALVE_FAULT.XV010_FAIL_TO_OPEN, FAIL_TO_CLOSE => "Valves Data".R10_VALVE_FAULT.XV10_FAIL_TO_CLOSE, status => "Valves Data".R10_XV10.STATUS)
   END_RUNG
   RUNG wire#powerrail
      Contact( "Valves Data".R10_XV10.RESET )
   END_RUNG wire#w1
   RUNG wire#powerrail
      Contact( "R10_DATA".R10.Reset )
   END_RUNG wire#w1
   RUNG wire#powerrail
      I_Contact( "DI_INPUTS".R10_INPUTS_RUA.EMG_PB )
   END_RUNG wire#w2
   // the same network as SCL:
   IF "AlwaysTRUE" THEN
       #valve_R10_XV10("auto/manual" := "Valves Data"."A/M".R10,   // "valve"
                       open_auto := "Valves Data".R10_XV10.CMD,
                       open_man := "Valves Data".R10_XV10.MCMD,
                       fbk_open := "A/GLR_010_XV401_OFB",
                       fbk_close := "A/GLR_010_XV401_CFB",
                       reset := "Valves Data".R10_XV10.RESET OR "R10_DATA".R10.Reset,
                       intl := NOT "DI_INPUTS".R10_INPUTS_RUA.EMG_PB,
                       Mon_En := 1,
                       mon_sp := "Valves Data".R10_XV10.MON_TIME,
                       SEMI := "Valves Data".SEMI_AUTO.R10,
                       "open/close" => "A/GLR_010_XV401_CMD",
                       FAIL_TO_OPEN => "Valves Data".R10_VALVE_FAULT.XV010_FAIL_TO_OPEN,
                       FAIL_TO_CLOSE => "Valves Data".R10_VALVE_FAULT.XV10_FAIL_TO_CLOSE,
                       status => "Valves Data".R10_XV10.STATUS);
   END_IF;
END_REGION

REGION Network 110: ****REACTOR_11****
END_REGION

REGION Network 111: R11_XV01
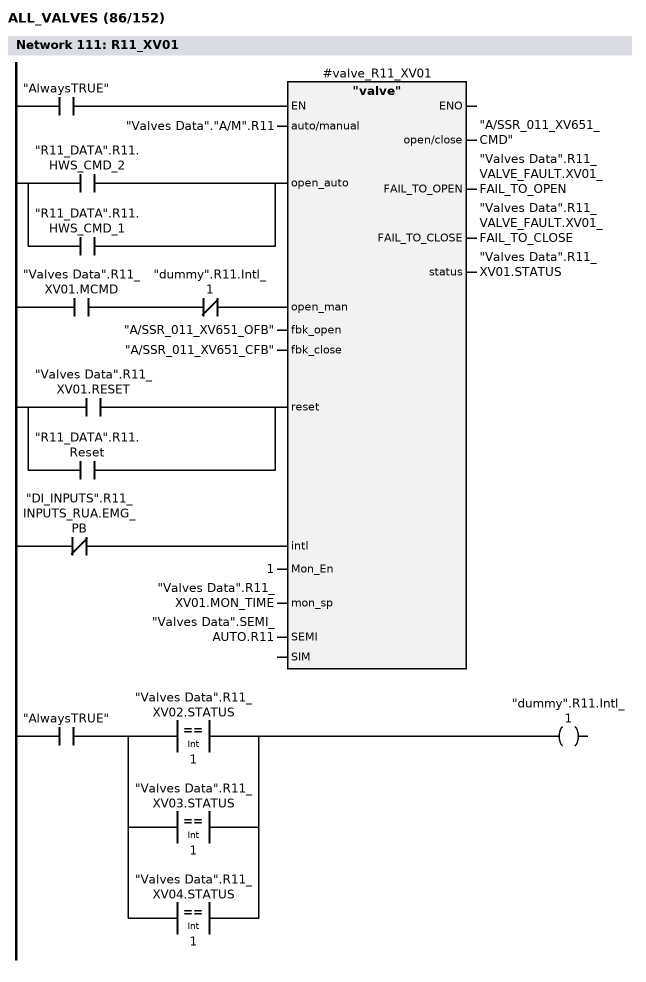
   RUNG wire#powerrail
      Contact( "AlwaysTRUE" )
      #valve_R11_XV01(open_auto := wire#w1, open_man := wire#w2, reset := wire#w3, intl := wire#w4, "auto/manual" := "Valves Data"."A/M".R11, fbk_open := "A/SSR_011_XV651_OFB", fbk_close := "A/SSR_011_XV651_CFB", Mon_En := 1, mon_sp := "Valves Data".R11_XV01.MON_TIME, SEMI := "Valves Data".SEMI_AUTO.R11, SIM :=, "open/close" => "A/SSR_011_XV651_CMD", FAIL_TO_OPEN => "Valves Data".R11_VALVE_FAULT.XV01_FAIL_TO_OPEN, FAIL_TO_CLOSE => "Valves Data".R11_VALVE_FAULT.XV01_FAIL_TO_CLOSE, status => "Valves Data".R11_XV01.STATUS)
   END_RUNG
   RUNG wire#powerrail
      Contact( "R11_DATA".R11.HWS_CMD_2 )
   END_RUNG wire#w1
   RUNG wire#powerrail
      Contact( "R11_DATA".R11.HWS_CMD_1 )
   END_RUNG wire#w1
   RUNG wire#powerrail
      Contact( "Valves Data".R11_XV01.MCMD )
      I_Contact( "dummy".R11.Intl_1 )
   END_RUNG wire#w2
   RUNG wire#powerrail
      Contact( "Valves Data".R11_XV01.RESET )
   END_RUNG wire#w3
   RUNG wire#powerrail
      Contact( "R11_DATA".R11.Reset )
   END_RUNG wire#w3
   RUNG wire#powerrail
      I_Contact( "DI_INPUTS".R11_INPUTS_RUA.EMG_PB )
   END_RUNG wire#w4
   RUNG wire#powerrail
      Contact( "AlwaysTRUE" )
      wire#w5
      { S7_Templates := "SrcType := Int" } EQ_Contact(in1 := "Valves Data".R11_XV02.STATUS, in2 := 1)
      wire#w6
      Coil( "dummy".R11.Intl_1 )
   END_RUNG
   RUNG wire#w5
      { S7_Templates := "SrcType := Int" } EQ_Contact(in1 := "Valves Data".R11_XV03.STATUS, in2 := 1)
   END_RUNG wire#w6
   RUNG wire#w5
      { S7_Templates := "SrcType := Int" } EQ_Contact(in1 := "Valves Data".R11_XV04.STATUS, in2 := 1)
   END_RUNG wire#w6
   // the same network as SCL:
   IF "AlwaysTRUE" THEN
       #valve_R11_XV01("auto/manual" := "Valves Data"."A/M".R11,   // "valve"
                       open_auto := "R11_DATA".R11.HWS_CMD_2 OR "R11_DATA".R11.HWS_CMD_1,
                       open_man := "Valves Data".R11_XV01.MCMD AND NOT "dummy".R11.Intl_1,
                       fbk_open := "A/SSR_011_XV651_OFB",
                       fbk_close := "A/SSR_011_XV651_CFB",
                       reset := "Valves Data".R11_XV01.RESET OR "R11_DATA".R11.Reset,
                       intl := NOT "DI_INPUTS".R11_INPUTS_RUA.EMG_PB,
                       Mon_En := 1,
                       mon_sp := "Valves Data".R11_XV01.MON_TIME,
                       SEMI := "Valves Data".SEMI_AUTO.R11,
                       "open/close" => "A/SSR_011_XV651_CMD",
                       FAIL_TO_OPEN => "Valves Data".R11_VALVE_FAULT.XV01_FAIL_TO_OPEN,
                       FAIL_TO_CLOSE => "Valves Data".R11_VALVE_FAULT.XV01_FAIL_TO_CLOSE,
                       status => "Valves Data".R11_XV01.STATUS);
   END_IF;
   "dummy".R11.Intl_1 := "AlwaysTRUE" AND (("Valves Data".R11_XV02.STATUS = 1) OR ("Valves Data".R11_XV03.STATUS = 1) OR ("Valves Data".R11_XV04.STATUS = 1));
END_REGION

REGION Network 112: R11_XV02
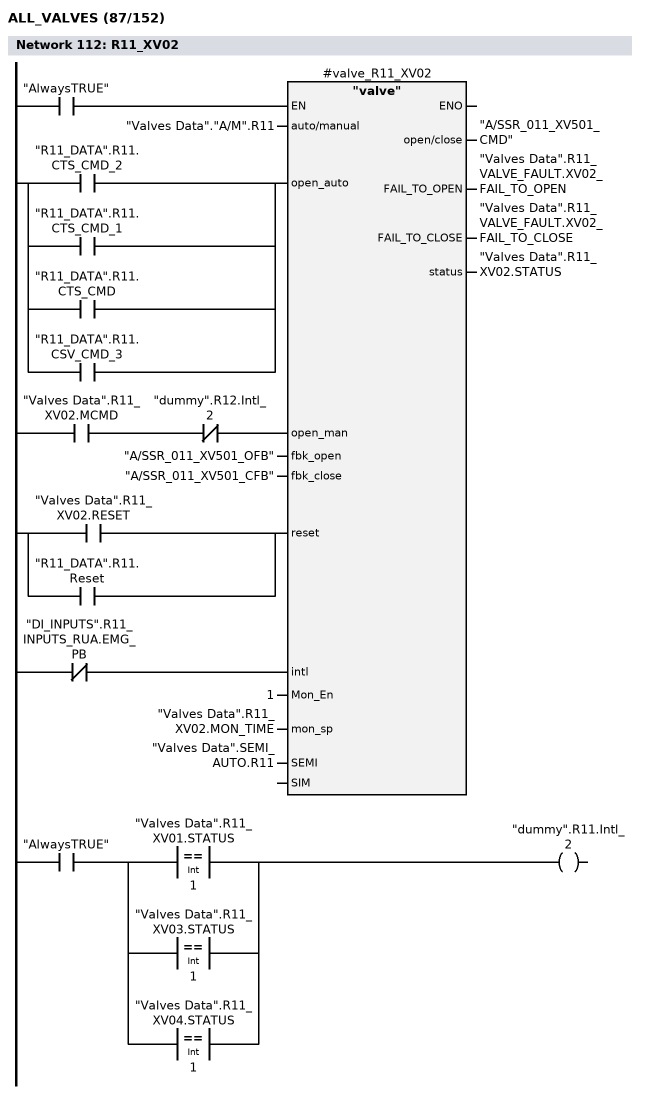
   RUNG wire#powerrail
      Contact( "AlwaysTRUE" )
      #valve_R11_XV02(open_auto := wire#w1, open_man := wire#w2, reset := wire#w3, intl := wire#w4, "auto/manual" := "Valves Data"."A/M".R11, fbk_open := "A/SSR_011_XV501_OFB", fbk_close := "A/SSR_011_XV501_CFB", Mon_En := 1, mon_sp := "Valves Data".R11_XV02.MON_TIME, SEMI := "Valves Data".SEMI_AUTO.R11, SIM :=, "open/close" => "A/SSR_011_XV501_CMD", FAIL_TO_OPEN => "Valves Data".R11_VALVE_FAULT.XV02_FAIL_TO_OPEN, FAIL_TO_CLOSE => "Valves Data".R11_VALVE_FAULT.XV02_FAIL_TO_CLOSE, status => "Valves Data".R11_XV02.STATUS)
   END_RUNG
   RUNG wire#powerrail
      Contact( "R11_DATA".R11.CTS_CMD_2 )
   END_RUNG wire#w1
   RUNG wire#powerrail
      Contact( "R11_DATA".R11.CTS_CMD_1 )
   END_RUNG wire#w1
   RUNG wire#powerrail
      Contact( "R11_DATA".R11.CTS_CMD )
   END_RUNG wire#w1
   RUNG wire#powerrail
      Contact( "R11_DATA".R11.CSV_CMD_3 )
   END_RUNG wire#w1
   RUNG wire#powerrail
      Contact( "Valves Data".R11_XV02.MCMD )
      I_Contact( "dummy".R12.Intl_2 )
   END_RUNG wire#w2
   RUNG wire#powerrail
      Contact( "Valves Data".R11_XV02.RESET )
   END_RUNG wire#w3
   RUNG wire#powerrail
      Contact( "R11_DATA".R11.Reset )
   END_RUNG wire#w3
   RUNG wire#powerrail
      I_Contact( "DI_INPUTS".R11_INPUTS_RUA.EMG_PB )
   END_RUNG wire#w4
   RUNG wire#powerrail
      Contact( "AlwaysTRUE" )
      wire#w5
      { S7_Templates := "SrcType := Int" } EQ_Contact(in1 := "Valves Data".R11_XV01.STATUS, in2 := 1)
      wire#w6
      Coil( "dummy".R11.Intl_2 )
   END_RUNG
   RUNG wire#w5
      { S7_Templates := "SrcType := Int" } EQ_Contact(in1 := "Valves Data".R11_XV03.STATUS, in2 := 1)
   END_RUNG wire#w6
   RUNG wire#w5
      { S7_Templates := "SrcType := Int" } EQ_Contact(in1 := "Valves Data".R11_XV04.STATUS, in2 := 1)
   END_RUNG wire#w6
   // the same network as SCL:
   IF "AlwaysTRUE" THEN
       #valve_R11_XV02("auto/manual" := "Valves Data"."A/M".R11,   // "valve"
                       open_auto := "R11_DATA".R11.CTS_CMD_2 OR "R11_DATA".R11.CTS_CMD_1 OR "R11_DATA".R11.CTS_CMD OR "R11_DATA".R11.CSV_CMD_3,
                       open_man := "Valves Data".R11_XV02.MCMD AND NOT "dummy".R12.Intl_2,
                       fbk_open := "A/SSR_011_XV501_OFB",
                       fbk_close := "A/SSR_011_XV501_CFB",
                       reset := "Valves Data".R11_XV02.RESET OR "R11_DATA".R11.Reset,
                       intl := NOT "DI_INPUTS".R11_INPUTS_RUA.EMG_PB,
                       Mon_En := 1,
                       mon_sp := "Valves Data".R11_XV02.MON_TIME,
                       SEMI := "Valves Data".SEMI_AUTO.R11,
                       "open/close" => "A/SSR_011_XV501_CMD",
                       FAIL_TO_OPEN => "Valves Data".R11_VALVE_FAULT.XV02_FAIL_TO_OPEN,
                       FAIL_TO_CLOSE => "Valves Data".R11_VALVE_FAULT.XV02_FAIL_TO_CLOSE,
                       status => "Valves Data".R11_XV02.STATUS);
   END_IF;
   "dummy".R11.Intl_2 := "AlwaysTRUE" AND (("Valves Data".R11_XV01.STATUS = 1) OR ("Valves Data".R11_XV03.STATUS = 1) OR ("Valves Data".R11_XV04.STATUS = 1));
END_REGION

REGION Network 113: R11_XV03
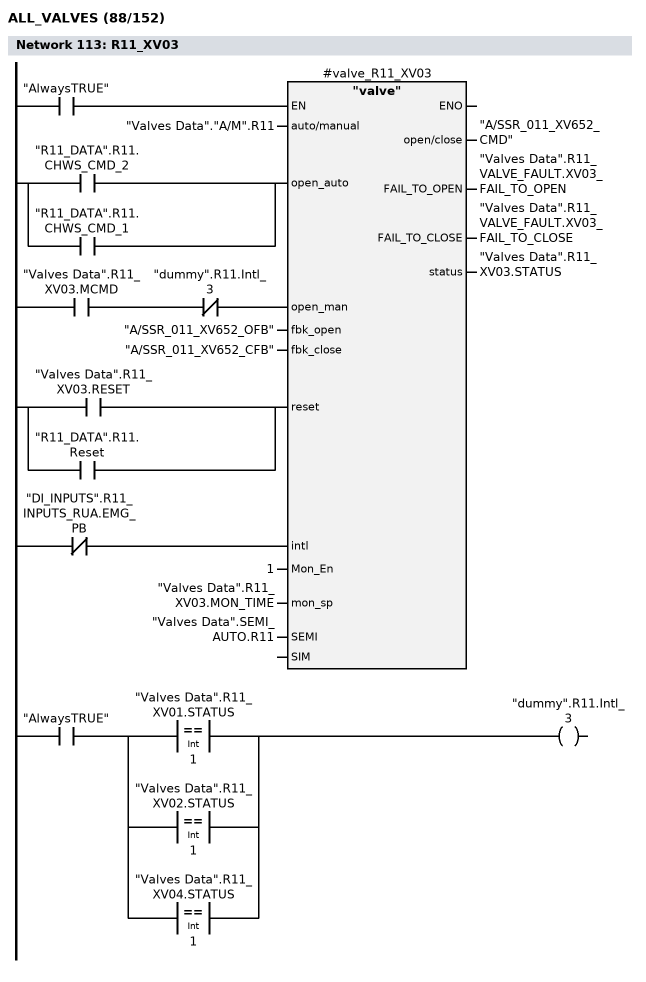
   RUNG wire#powerrail
      Contact( "AlwaysTRUE" )
      #valve_R11_XV03(open_auto := wire#w1, open_man := wire#w2, reset := wire#w3, intl := wire#w4, "auto/manual" := "Valves Data"."A/M".R11, fbk_open := "A/SSR_011_XV652_OFB", fbk_close := "A/SSR_011_XV652_CFB", Mon_En := 1, mon_sp := "Valves Data".R11_XV03.MON_TIME, SEMI := "Valves Data".SEMI_AUTO.R11, SIM :=, "open/close" => "A/SSR_011_XV652_CMD", FAIL_TO_OPEN => "Valves Data".R11_VALVE_FAULT.XV03_FAIL_TO_OPEN, FAIL_TO_CLOSE => "Valves Data".R11_VALVE_FAULT.XV03_FAIL_TO_CLOSE, status => "Valves Data".R11_XV03.STATUS)
   END_RUNG
   RUNG wire#powerrail
      Contact( "R11_DATA".R11.CHWS_CMD_2 )
   END_RUNG wire#w1
   RUNG wire#powerrail
      Contact( "R11_DATA".R11.CHWS_CMD_1 )
   END_RUNG wire#w1
   RUNG wire#powerrail
      Contact( "Valves Data".R11_XV03.MCMD )
      I_Contact( "dummy".R11.Intl_3 )
   END_RUNG wire#w2
   RUNG wire#powerrail
      Contact( "Valves Data".R11_XV03.RESET )
   END_RUNG wire#w3
   RUNG wire#powerrail
      Contact( "R11_DATA".R11.Reset )
   END_RUNG wire#w3
   RUNG wire#powerrail
      I_Contact( "DI_INPUTS".R11_INPUTS_RUA.EMG_PB )
   END_RUNG wire#w4
   RUNG wire#powerrail
      Contact( "AlwaysTRUE" )
      wire#w5
      { S7_Templates := "SrcType := Int" } EQ_Contact(in1 := "Valves Data".R11_XV01.STATUS, in2 := 1)
      wire#w6
      Coil( "dummy".R11.Intl_3 )
   END_RUNG
   RUNG wire#w5
      { S7_Templates := "SrcType := Int" } EQ_Contact(in1 := "Valves Data".R11_XV02.STATUS, in2 := 1)
   END_RUNG wire#w6
   RUNG wire#w5
      { S7_Templates := "SrcType := Int" } EQ_Contact(in1 := "Valves Data".R11_XV04.STATUS, in2 := 1)
   END_RUNG wire#w6
   // the same network as SCL:
   IF "AlwaysTRUE" THEN
       #valve_R11_XV03("auto/manual" := "Valves Data"."A/M".R11,   // "valve"
                       open_auto := "R11_DATA".R11.CHWS_CMD_2 OR "R11_DATA".R11.CHWS_CMD_1,
                       open_man := "Valves Data".R11_XV03.MCMD AND NOT "dummy".R11.Intl_3,
                       fbk_open := "A/SSR_011_XV652_OFB",
                       fbk_close := "A/SSR_011_XV652_CFB",
                       reset := "Valves Data".R11_XV03.RESET OR "R11_DATA".R11.Reset,
                       intl := NOT "DI_INPUTS".R11_INPUTS_RUA.EMG_PB,
                       Mon_En := 1,
                       mon_sp := "Valves Data".R11_XV03.MON_TIME,
                       SEMI := "Valves Data".SEMI_AUTO.R11,
                       "open/close" => "A/SSR_011_XV652_CMD",
                       FAIL_TO_OPEN => "Valves Data".R11_VALVE_FAULT.XV03_FAIL_TO_OPEN,
                       FAIL_TO_CLOSE => "Valves Data".R11_VALVE_FAULT.XV03_FAIL_TO_CLOSE,
                       status => "Valves Data".R11_XV03.STATUS);
   END_IF;
   "dummy".R11.Intl_3 := "AlwaysTRUE" AND (("Valves Data".R11_XV01.STATUS = 1) OR ("Valves Data".R11_XV02.STATUS = 1) OR ("Valves Data".R11_XV04.STATUS = 1));
END_REGION

REGION Network 114: R11_XV04
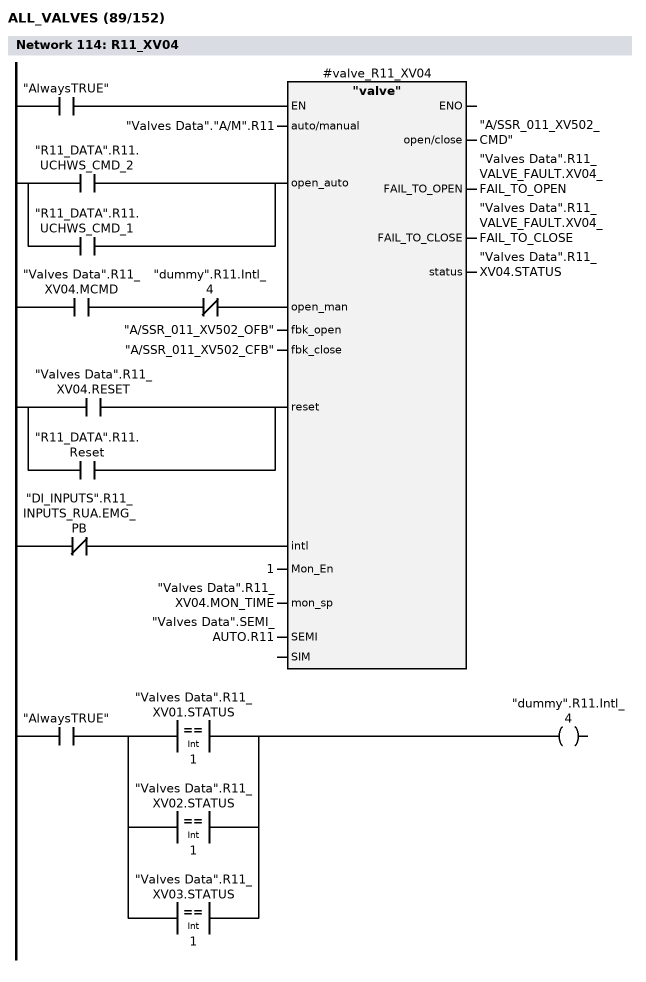
   RUNG wire#powerrail
      Contact( "AlwaysTRUE" )
      #valve_R11_XV04(open_auto := wire#w1, open_man := wire#w2, reset := wire#w3, intl := wire#w4, "auto/manual" := "Valves Data"."A/M".R11, fbk_open := "A/SSR_011_XV502_OFB", fbk_close := "A/SSR_011_XV502_CFB", Mon_En := 1, mon_sp := "Valves Data".R11_XV04.MON_TIME, SEMI := "Valves Data".SEMI_AUTO.R11, SIM :=, "open/close" => "A/SSR_011_XV502_CMD", FAIL_TO_OPEN => "Valves Data".R11_VALVE_FAULT.XV04_FAIL_TO_OPEN, FAIL_TO_CLOSE => "Valves Data".R11_VALVE_FAULT.XV04_FAIL_TO_CLOSE, status => "Valves Data".R11_XV04.STATUS)
   END_RUNG
   RUNG wire#powerrail
      Contact( "R11_DATA".R11.UCHWS_CMD_2 )
   END_RUNG wire#w1
   RUNG wire#powerrail
      Contact( "R11_DATA".R11.UCHWS_CMD_1 )
   END_RUNG wire#w1
   RUNG wire#powerrail
      Contact( "Valves Data".R11_XV04.MCMD )
      I_Contact( "dummy".R11.Intl_4 )
   END_RUNG wire#w2
   RUNG wire#powerrail
      Contact( "Valves Data".R11_XV04.RESET )
   END_RUNG wire#w3
   RUNG wire#powerrail
      Contact( "R11_DATA".R11.Reset )
   END_RUNG wire#w3
   RUNG wire#powerrail
      I_Contact( "DI_INPUTS".R11_INPUTS_RUA.EMG_PB )
   END_RUNG wire#w4
   RUNG wire#powerrail
      Contact( "AlwaysTRUE" )
      wire#w5
      { S7_Templates := "SrcType := Int" } EQ_Contact(in1 := "Valves Data".R11_XV01.STATUS, in2 := 1)
      wire#w6
      Coil( "dummy".R11.Intl_4 )
   END_RUNG
   RUNG wire#w5
      { S7_Templates := "SrcType := Int" } EQ_Contact(in1 := "Valves Data".R11_XV02.STATUS, in2 := 1)
   END_RUNG wire#w6
   RUNG wire#w5
      { S7_Templates := "SrcType := Int" } EQ_Contact(in1 := "Valves Data".R11_XV03.STATUS, in2 := 1)
   END_RUNG wire#w6
   // the same network as SCL:
   IF "AlwaysTRUE" THEN
       #valve_R11_XV04("auto/manual" := "Valves Data"."A/M".R11,   // "valve"
                       open_auto := "R11_DATA".R11.UCHWS_CMD_2 OR "R11_DATA".R11.UCHWS_CMD_1,
                       open_man := "Valves Data".R11_XV04.MCMD AND NOT "dummy".R11.Intl_4,
                       fbk_open := "A/SSR_011_XV502_OFB",
                       fbk_close := "A/SSR_011_XV502_CFB",
                       reset := "Valves Data".R11_XV04.RESET OR "R11_DATA".R11.Reset,
                       intl := NOT "DI_INPUTS".R11_INPUTS_RUA.EMG_PB,
                       Mon_En := 1,
                       mon_sp := "Valves Data".R11_XV04.MON_TIME,
                       SEMI := "Valves Data".SEMI_AUTO.R11,
                       "open/close" => "A/SSR_011_XV502_CMD",
                       FAIL_TO_OPEN => "Valves Data".R11_VALVE_FAULT.XV04_FAIL_TO_OPEN,
                       FAIL_TO_CLOSE => "Valves Data".R11_VALVE_FAULT.XV04_FAIL_TO_CLOSE,
                       status => "Valves Data".R11_XV04.STATUS);
   END_IF;
   "dummy".R11.Intl_4 := "AlwaysTRUE" AND (("Valves Data".R11_XV01.STATUS = 1) OR ("Valves Data".R11_XV02.STATUS = 1) OR ("Valves Data".R11_XV03.STATUS = 1));
END_REGION

REGION Network 115: R11_XV05
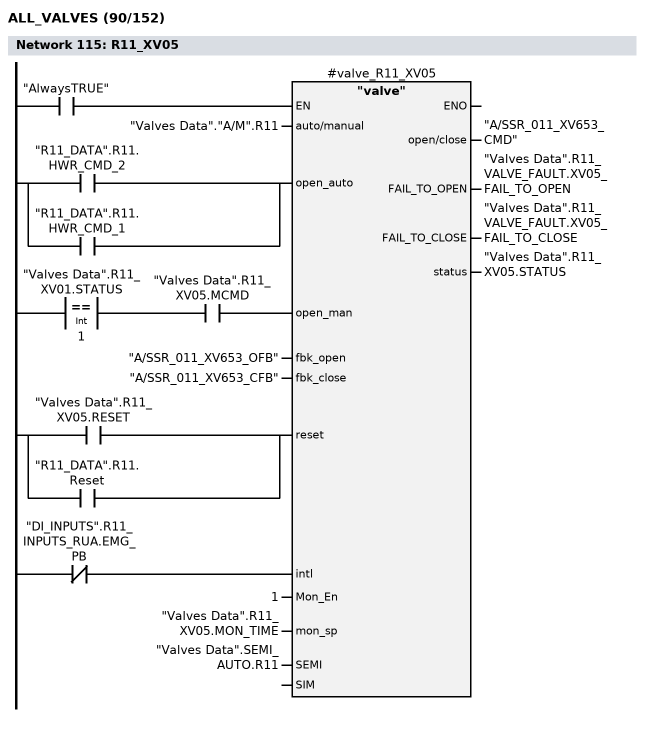
   RUNG wire#powerrail
      Contact( "AlwaysTRUE" )
      #valve_R11_XV05(open_auto := wire#w1, open_man := wire#w2, reset := wire#w3, intl := wire#w4, "auto/manual" := "Valves Data"."A/M".R11, fbk_open := "A/SSR_011_XV653_OFB", fbk_close := "A/SSR_011_XV653_CFB", Mon_En := 1, mon_sp := "Valves Data".R11_XV05.MON_TIME, SEMI := "Valves Data".SEMI_AUTO.R11, SIM :=, "open/close" => "A/SSR_011_XV653_CMD", FAIL_TO_OPEN => "Valves Data".R11_VALVE_FAULT.XV05_FAIL_TO_OPEN, FAIL_TO_CLOSE => "Valves Data".R11_VALVE_FAULT.XV05_FAIL_TO_CLOSE, status => "Valves Data".R11_XV05.STATUS)
   END_RUNG
   RUNG wire#powerrail
      Contact( "R11_DATA".R11.HWR_CMD_2 )
   END_RUNG wire#w1
   RUNG wire#powerrail
      Contact( "R11_DATA".R11.HWR_CMD_1 )
   END_RUNG wire#w1
   RUNG wire#powerrail
      { S7_Templates := "SrcType := Int" } EQ_Contact(in1 := "Valves Data".R11_XV01.STATUS, in2 := 1)
      Contact( "Valves Data".R11_XV05.MCMD )
   END_RUNG wire#w2
   RUNG wire#powerrail
      Contact( "Valves Data".R11_XV05.RESET )
   END_RUNG wire#w3
   RUNG wire#powerrail
      Contact( "R11_DATA".R11.Reset )
   END_RUNG wire#w3
   RUNG wire#powerrail
      I_Contact( "DI_INPUTS".R11_INPUTS_RUA.EMG_PB )
   END_RUNG wire#w4
   // the same network as SCL:
   IF "AlwaysTRUE" THEN
       #valve_R11_XV05("auto/manual" := "Valves Data"."A/M".R11,   // "valve"
                       open_auto := "R11_DATA".R11.HWR_CMD_2 OR "R11_DATA".R11.HWR_CMD_1,
                       open_man := ("Valves Data".R11_XV01.STATUS = 1) AND "Valves Data".R11_XV05.MCMD,
                       fbk_open := "A/SSR_011_XV653_OFB",
                       fbk_close := "A/SSR_011_XV653_CFB",
                       reset := "Valves Data".R11_XV05.RESET OR "R11_DATA".R11.Reset,
                       intl := NOT "DI_INPUTS".R11_INPUTS_RUA.EMG_PB,
                       Mon_En := 1,
                       mon_sp := "Valves Data".R11_XV05.MON_TIME,
                       SEMI := "Valves Data".SEMI_AUTO.R11,
                       "open/close" => "A/SSR_011_XV653_CMD",
                       FAIL_TO_OPEN => "Valves Data".R11_VALVE_FAULT.XV05_FAIL_TO_OPEN,
                       FAIL_TO_CLOSE => "Valves Data".R11_VALVE_FAULT.XV05_FAIL_TO_CLOSE,
                       status => "Valves Data".R11_XV05.STATUS);
   END_IF;
END_REGION

REGION Network 116: R11_XV06
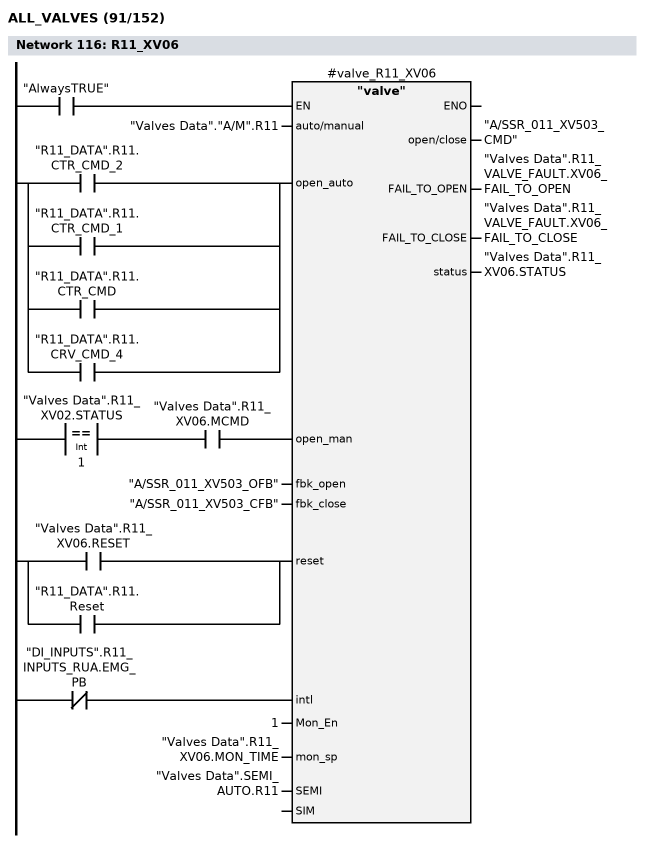
   RUNG wire#powerrail
      Contact( "AlwaysTRUE" )
      #valve_R11_XV06(open_auto := wire#w1, open_man := wire#w2, reset := wire#w3, intl := wire#w4, "auto/manual" := "Valves Data"."A/M".R11, fbk_open := "A/SSR_011_XV503_OFB", fbk_close := "A/SSR_011_XV503_CFB", Mon_En := 1, mon_sp := "Valves Data".R11_XV06.MON_TIME, SEMI := "Valves Data".SEMI_AUTO.R11, SIM :=, "open/close" => "A/SSR_011_XV503_CMD", FAIL_TO_OPEN => "Valves Data".R11_VALVE_FAULT.XV06_FAIL_TO_OPEN, FAIL_TO_CLOSE => "Valves Data".R11_VALVE_FAULT.XV06_FAIL_TO_CLOSE, status => "Valves Data".R11_XV06.STATUS)
   END_RUNG
   RUNG wire#powerrail
      Contact( "R11_DATA".R11.CTR_CMD_2 )
   END_RUNG wire#w1
   RUNG wire#powerrail
      Contact( "R11_DATA".R11.CTR_CMD_1 )
   END_RUNG wire#w1
   RUNG wire#powerrail
      Contact( "R11_DATA".R11.CTR_CMD )
   END_RUNG wire#w1
   RUNG wire#powerrail
      Contact( "R11_DATA".R11.CRV_CMD_4 )
   END_RUNG wire#w1
   RUNG wire#powerrail
      { S7_Templates := "SrcType := Int" } EQ_Contact(in1 := "Valves Data".R11_XV02.STATUS, in2 := 1)
      Contact( "Valves Data".R11_XV06.MCMD )
   END_RUNG wire#w2
   RUNG wire#powerrail
      Contact( "Valves Data".R11_XV06.RESET )
   END_RUNG wire#w3
   RUNG wire#powerrail
      Contact( "R11_DATA".R11.Reset )
   END_RUNG wire#w3
   RUNG wire#powerrail
      I_Contact( "DI_INPUTS".R11_INPUTS_RUA.EMG_PB )
   END_RUNG wire#w4
   // the same network as SCL:
   IF "AlwaysTRUE" THEN
       #valve_R11_XV06("auto/manual" := "Valves Data"."A/M".R11,   // "valve"
                       open_auto := "R11_DATA".R11.CTR_CMD_2 OR "R11_DATA".R11.CTR_CMD_1 OR "R11_DATA".R11.CTR_CMD OR "R11_DATA".R11.CRV_CMD_4,
                       open_man := ("Valves Data".R11_XV02.STATUS = 1) AND "Valves Data".R11_XV06.MCMD,
                       fbk_open := "A/SSR_011_XV503_OFB",
                       fbk_close := "A/SSR_011_XV503_CFB",
                       reset := "Valves Data".R11_XV06.RESET OR "R11_DATA".R11.Reset,
                       intl := NOT "DI_INPUTS".R11_INPUTS_RUA.EMG_PB,
                       Mon_En := 1,
                       mon_sp := "Valves Data".R11_XV06.MON_TIME,
                       SEMI := "Valves Data".SEMI_AUTO.R11,
                       "open/close" => "A/SSR_011_XV503_CMD",
                       FAIL_TO_OPEN => "Valves Data".R11_VALVE_FAULT.XV06_FAIL_TO_OPEN,
                       FAIL_TO_CLOSE => "Valves Data".R11_VALVE_FAULT.XV06_FAIL_TO_CLOSE,
                       status => "Valves Data".R11_XV06.STATUS);
   END_IF;
END_REGION

REGION Network 117: R11_XV07
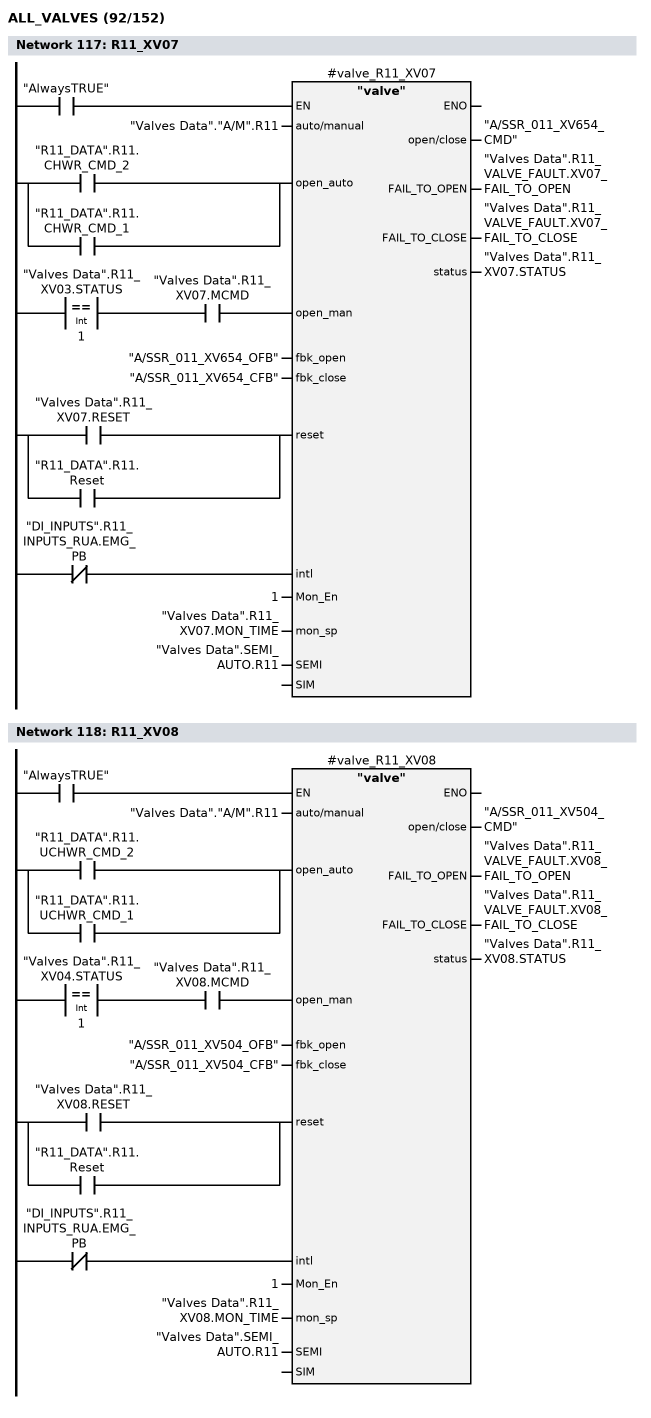
   RUNG wire#powerrail
      Contact( "AlwaysTRUE" )
      #valve_R11_XV07(open_auto := wire#w1, open_man := wire#w2, reset := wire#w3, intl := wire#w4, "auto/manual" := "Valves Data"."A/M".R11, fbk_open := "A/SSR_011_XV654_OFB", fbk_close := "A/SSR_011_XV654_CFB", Mon_En := 1, mon_sp := "Valves Data".R11_XV07.MON_TIME, SEMI := "Valves Data".SEMI_AUTO.R11, SIM :=, "open/close" => "A/SSR_011_XV654_CMD", FAIL_TO_OPEN => "Valves Data".R11_VALVE_FAULT.XV07_FAIL_TO_OPEN, FAIL_TO_CLOSE => "Valves Data".R11_VALVE_FAULT.XV07_FAIL_TO_CLOSE, status => "Valves Data".R11_XV07.STATUS)
   END_RUNG
   RUNG wire#powerrail
      Contact( "R11_DATA".R11.CHWR_CMD_2 )
   END_RUNG wire#w1
   RUNG wire#powerrail
      Contact( "R11_DATA".R11.CHWR_CMD_1 )
   END_RUNG wire#w1
   RUNG wire#powerrail
      { S7_Templates := "SrcType := Int" } EQ_Contact(in1 := "Valves Data".R11_XV03.STATUS, in2 := 1)
      Contact( "Valves Data".R11_XV07.MCMD )
   END_RUNG wire#w2
   RUNG wire#powerrail
      Contact( "Valves Data".R11_XV07.RESET )
   END_RUNG wire#w3
   RUNG wire#powerrail
      Contact( "R11_DATA".R11.Reset )
   END_RUNG wire#w3
   RUNG wire#powerrail
      I_Contact( "DI_INPUTS".R11_INPUTS_RUA.EMG_PB )
   END_RUNG wire#w4
   // the same network as SCL:
   IF "AlwaysTRUE" THEN
       #valve_R11_XV07("auto/manual" := "Valves Data"."A/M".R11,   // "valve"
                       open_auto := "R11_DATA".R11.CHWR_CMD_2 OR "R11_DATA".R11.CHWR_CMD_1,
                       open_man := ("Valves Data".R11_XV03.STATUS = 1) AND "Valves Data".R11_XV07.MCMD,
                       fbk_open := "A/SSR_011_XV654_OFB",
                       fbk_close := "A/SSR_011_XV654_CFB",
                       reset := "Valves Data".R11_XV07.RESET OR "R11_DATA".R11.Reset,
                       intl := NOT "DI_INPUTS".R11_INPUTS_RUA.EMG_PB,
                       Mon_En := 1,
                       mon_sp := "Valves Data".R11_XV07.MON_TIME,
                       SEMI := "Valves Data".SEMI_AUTO.R11,
                       "open/close" => "A/SSR_011_XV654_CMD",
                       FAIL_TO_OPEN => "Valves Data".R11_VALVE_FAULT.XV07_FAIL_TO_OPEN,
                       FAIL_TO_CLOSE => "Valves Data".R11_VALVE_FAULT.XV07_FAIL_TO_CLOSE,
                       status => "Valves Data".R11_XV07.STATUS);
   END_IF;
END_REGION

REGION Network 118: R11_XV08
   RUNG wire#powerrail
      Contact( "AlwaysTRUE" )
      #valve_R11_XV08(open_auto := wire#w1, open_man := wire#w2, reset := wire#w3, intl := wire#w4, "auto/manual" := "Valves Data"."A/M".R11, fbk_open := "A/SSR_011_XV504_OFB", fbk_close := "A/SSR_011_XV504_CFB", Mon_En := 1, mon_sp := "Valves Data".R11_XV08.MON_TIME, SEMI := "Valves Data".SEMI_AUTO.R11, SIM :=, "open/close" => "A/SSR_011_XV504_CMD", FAIL_TO_OPEN => "Valves Data".R11_VALVE_FAULT.XV08_FAIL_TO_OPEN, FAIL_TO_CLOSE => "Valves Data".R11_VALVE_FAULT.XV08_FAIL_TO_CLOSE, status => "Valves Data".R11_XV08.STATUS)
   END_RUNG
   RUNG wire#powerrail
      Contact( "R11_DATA".R11.UCHWR_CMD_2 )
   END_RUNG wire#w1
   RUNG wire#powerrail
      Contact( "R11_DATA".R11.UCHWR_CMD_1 )
   END_RUNG wire#w1
   RUNG wire#powerrail
      { S7_Templates := "SrcType := Int" } EQ_Contact(in1 := "Valves Data".R11_XV04.STATUS, in2 := 1)
      Contact( "Valves Data".R11_XV08.MCMD )
   END_RUNG wire#w2
   RUNG wire#powerrail
      Contact( "Valves Data".R11_XV08.RESET )
   END_RUNG wire#w3
   RUNG wire#powerrail
      Contact( "R11_DATA".R11.Reset )
   END_RUNG wire#w3
   RUNG wire#powerrail
      I_Contact( "DI_INPUTS".R11_INPUTS_RUA.EMG_PB )
   END_RUNG wire#w4
   // the same network as SCL:
   IF "AlwaysTRUE" THEN
       #valve_R11_XV08("auto/manual" := "Valves Data"."A/M".R11,   // "valve"
                       open_auto := "R11_DATA".R11.UCHWR_CMD_2 OR "R11_DATA".R11.UCHWR_CMD_1,
                       open_man := ("Valves Data".R11_XV04.STATUS = 1) AND "Valves Data".R11_XV08.MCMD,
                       fbk_open := "A/SSR_011_XV504_OFB",
                       fbk_close := "A/SSR_011_XV504_CFB",
                       reset := "Valves Data".R11_XV08.RESET OR "R11_DATA".R11.Reset,
                       intl := NOT "DI_INPUTS".R11_INPUTS_RUA.EMG_PB,
                       Mon_En := 1,
                       mon_sp := "Valves Data".R11_XV08.MON_TIME,
                       SEMI := "Valves Data".SEMI_AUTO.R11,
                       "open/close" => "A/SSR_011_XV504_CMD",
                       FAIL_TO_OPEN => "Valves Data".R11_VALVE_FAULT.XV08_FAIL_TO_OPEN,
                       FAIL_TO_CLOSE => "Valves Data".R11_VALVE_FAULT.XV08_FAIL_TO_CLOSE,
                       status => "Valves Data".R11_XV08.STATUS);
   END_IF;
END_REGION

REGION Network 119: R11_XV09
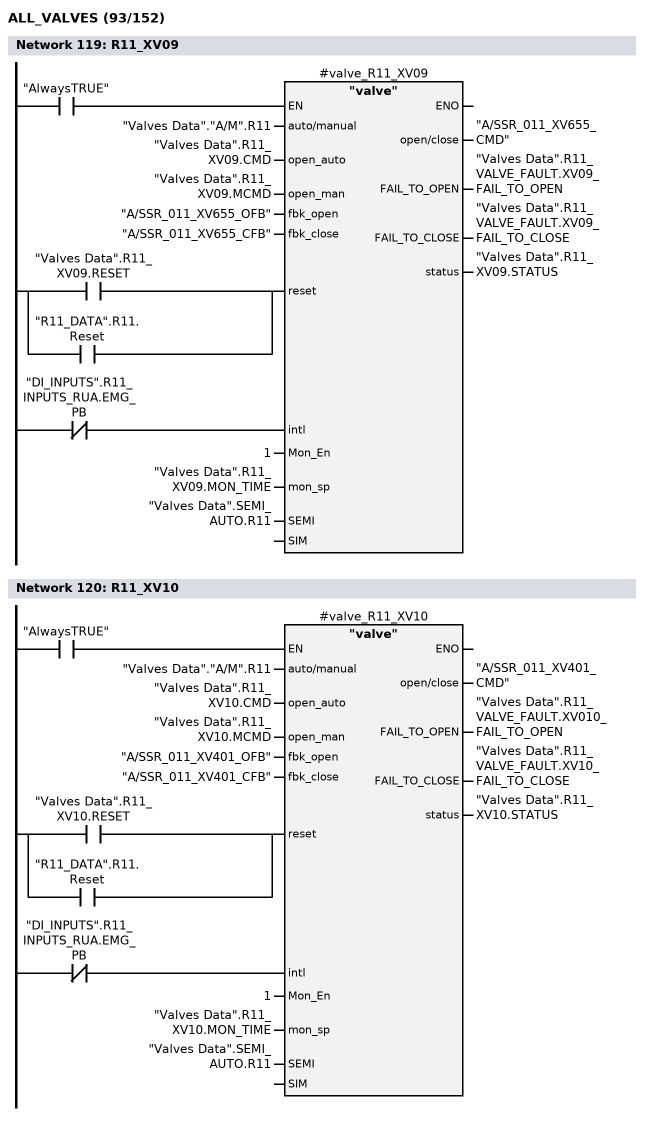
   RUNG wire#powerrail
      Contact( "AlwaysTRUE" )
      #valve_R11_XV09(reset := wire#w1, intl := wire#w2, "auto/manual" := "Valves Data"."A/M".R11, open_auto := "Valves Data".R11_XV09.CMD, open_man := "Valves Data".R11_XV09.MCMD, fbk_open := "A/SSR_011_XV655_OFB", fbk_close := "A/SSR_011_XV655_CFB", Mon_En := 1, mon_sp := "Valves Data".R11_XV09.MON_TIME, SEMI := "Valves Data".SEMI_AUTO.R11, SIM :=, "open/close" => "A/SSR_011_XV655_CMD", FAIL_TO_OPEN => "Valves Data".R11_VALVE_FAULT.XV09_FAIL_TO_OPEN, FAIL_TO_CLOSE => "Valves Data".R11_VALVE_FAULT.XV09_FAIL_TO_CLOSE, status => "Valves Data".R11_XV09.STATUS)
   END_RUNG
   RUNG wire#powerrail
      Contact( "Valves Data".R11_XV09.RESET )
   END_RUNG wire#w1
   RUNG wire#powerrail
      Contact( "R11_DATA".R11.Reset )
   END_RUNG wire#w1
   RUNG wire#powerrail
      I_Contact( "DI_INPUTS".R11_INPUTS_RUA.EMG_PB )
   END_RUNG wire#w2
   // the same network as SCL:
   IF "AlwaysTRUE" THEN
       #valve_R11_XV09("auto/manual" := "Valves Data"."A/M".R11,   // "valve"
                       open_auto := "Valves Data".R11_XV09.CMD,
                       open_man := "Valves Data".R11_XV09.MCMD,
                       fbk_open := "A/SSR_011_XV655_OFB",
                       fbk_close := "A/SSR_011_XV655_CFB",
                       reset := "Valves Data".R11_XV09.RESET OR "R11_DATA".R11.Reset,
                       intl := NOT "DI_INPUTS".R11_INPUTS_RUA.EMG_PB,
                       Mon_En := 1,
                       mon_sp := "Valves Data".R11_XV09.MON_TIME,
                       SEMI := "Valves Data".SEMI_AUTO.R11,
                       "open/close" => "A/SSR_011_XV655_CMD",
                       FAIL_TO_OPEN => "Valves Data".R11_VALVE_FAULT.XV09_FAIL_TO_OPEN,
                       FAIL_TO_CLOSE => "Valves Data".R11_VALVE_FAULT.XV09_FAIL_TO_CLOSE,
                       status => "Valves Data".R11_XV09.STATUS);
   END_IF;
END_REGION

REGION Network 120: R11_XV10
   RUNG wire#powerrail
      Contact( "AlwaysTRUE" )
      #valve_R11_XV10(reset := wire#w1, intl := wire#w2, "auto/manual" := "Valves Data"."A/M".R11, open_auto := "Valves Data".R11_XV10.CMD, open_man := "Valves Data".R11_XV10.MCMD, fbk_open := "A/SSR_011_XV401_OFB", fbk_close := "A/SSR_011_XV401_CFB", Mon_En := 1, mon_sp := "Valves Data".R11_XV10.MON_TIME, SEMI := "Valves Data".SEMI_AUTO.R11, SIM :=, "open/close" => "A/SSR_011_XV401_CMD", FAIL_TO_OPEN => "Valves Data".R11_VALVE_FAULT.XV010_FAIL_TO_OPEN, FAIL_TO_CLOSE => "Valves Data".R11_VALVE_FAULT.XV10_FAIL_TO_CLOSE, status => "Valves Data".R11_XV10.STATUS)
   END_RUNG
   RUNG wire#powerrail
      Contact( "Valves Data".R11_XV10.RESET )
   END_RUNG wire#w1
   RUNG wire#powerrail
      Contact( "R11_DATA".R11.Reset )
   END_RUNG wire#w1
   RUNG wire#powerrail
      I_Contact( "DI_INPUTS".R11_INPUTS_RUA.EMG_PB )
   END_RUNG wire#w2
   // the same network as SCL:
   IF "AlwaysTRUE" THEN
       #valve_R11_XV10("auto/manual" := "Valves Data"."A/M".R11,   // "valve"
                       open_auto := "Valves Data".R11_XV10.CMD,
                       open_man := "Valves Data".R11_XV10.MCMD,
                       fbk_open := "A/SSR_011_XV401_OFB",
                       fbk_close := "A/SSR_011_XV401_CFB",
                       reset := "Valves Data".R11_XV10.RESET OR "R11_DATA".R11.Reset,
                       intl := NOT "DI_INPUTS".R11_INPUTS_RUA.EMG_PB,
                       Mon_En := 1,
                       mon_sp := "Valves Data".R11_XV10.MON_TIME,
                       SEMI := "Valves Data".SEMI_AUTO.R11,
                       "open/close" => "A/SSR_011_XV401_CMD",
                       FAIL_TO_OPEN => "Valves Data".R11_VALVE_FAULT.XV010_FAIL_TO_OPEN,
                       FAIL_TO_CLOSE => "Valves Data".R11_VALVE_FAULT.XV10_FAIL_TO_CLOSE,
                       status => "Valves Data".R11_XV10.STATUS);
   END_IF;
END_REGION

REGION Network 121: ****REACTOR_12****
END_REGION

REGION Network 122: R12_XV01
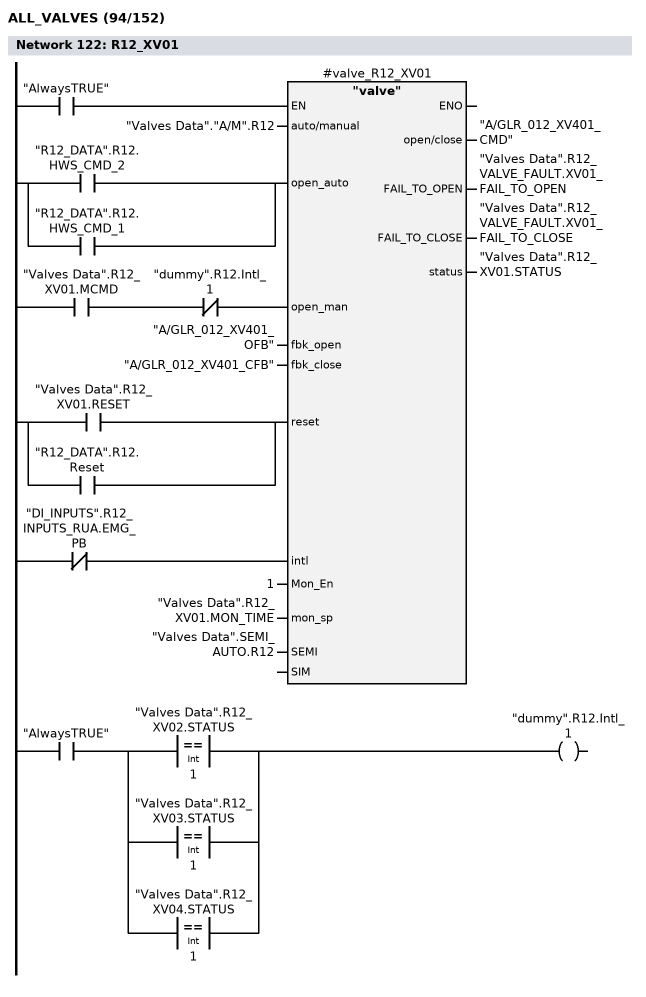
   RUNG wire#powerrail
      Contact( "AlwaysTRUE" )
      #valve_R12_XV01(open_auto := wire#w1, open_man := wire#w2, reset := wire#w3, intl := wire#w4, "auto/manual" := "Valves Data"."A/M".R12, fbk_open := "A/GLR_012_XV401_OFB", fbk_close := "A/GLR_012_XV401_CFB", Mon_En := 1, mon_sp := "Valves Data".R12_XV01.MON_TIME, SEMI := "Valves Data".SEMI_AUTO.R12, SIM :=, "open/close" => "A/GLR_012_XV401_CMD", FAIL_TO_OPEN => "Valves Data".R12_VALVE_FAULT.XV01_FAIL_TO_OPEN, FAIL_TO_CLOSE => "Valves Data".R12_VALVE_FAULT.XV01_FAIL_TO_CLOSE, status => "Valves Data".R12_XV01.STATUS)
   END_RUNG
   RUNG wire#powerrail
      Contact( "R12_DATA".R12.HWS_CMD_2 )
   END_RUNG wire#w1
   RUNG wire#powerrail
      Contact( "R12_DATA".R12.HWS_CMD_1 )
   END_RUNG wire#w1
   RUNG wire#powerrail
      Contact( "Valves Data".R12_XV01.MCMD )
      I_Contact( "dummy".R12.Intl_1 )
   END_RUNG wire#w2
   RUNG wire#powerrail
      Contact( "Valves Data".R12_XV01.RESET )
   END_RUNG wire#w3
   RUNG wire#powerrail
      Contact( "R12_DATA".R12.Reset )
   END_RUNG wire#w3
   RUNG wire#powerrail
      I_Contact( "DI_INPUTS".R12_INPUTS_RUA.EMG_PB )
   END_RUNG wire#w4
   RUNG wire#powerrail
      Contact( "AlwaysTRUE" )
      wire#w5
      { S7_Templates := "SrcType := Int" } EQ_Contact(in1 := "Valves Data".R12_XV02.STATUS, in2 := 1)
      wire#w6
      Coil( "dummy".R12.Intl_1 )
   END_RUNG
   RUNG wire#w5
      { S7_Templates := "SrcType := Int" } EQ_Contact(in1 := "Valves Data".R12_XV03.STATUS, in2 := 1)
   END_RUNG wire#w6
   RUNG wire#w5
      { S7_Templates := "SrcType := Int" } EQ_Contact(in1 := "Valves Data".R12_XV04.STATUS, in2 := 1)
   END_RUNG wire#w6
   // the same network as SCL:
   IF "AlwaysTRUE" THEN
       #valve_R12_XV01("auto/manual" := "Valves Data"."A/M".R12,   // "valve"
                       open_auto := "R12_DATA".R12.HWS_CMD_2 OR "R12_DATA".R12.HWS_CMD_1,
                       open_man := "Valves Data".R12_XV01.MCMD AND NOT "dummy".R12.Intl_1,
                       fbk_open := "A/GLR_012_XV401_OFB",
                       fbk_close := "A/GLR_012_XV401_CFB",
                       reset := "Valves Data".R12_XV01.RESET OR "R12_DATA".R12.Reset,
                       intl := NOT "DI_INPUTS".R12_INPUTS_RUA.EMG_PB,
                       Mon_En := 1,
                       mon_sp := "Valves Data".R12_XV01.MON_TIME,
                       SEMI := "Valves Data".SEMI_AUTO.R12,
                       "open/close" => "A/GLR_012_XV401_CMD",
                       FAIL_TO_OPEN => "Valves Data".R12_VALVE_FAULT.XV01_FAIL_TO_OPEN,
                       FAIL_TO_CLOSE => "Valves Data".R12_VALVE_FAULT.XV01_FAIL_TO_CLOSE,
                       status => "Valves Data".R12_XV01.STATUS);
   END_IF;
   "dummy".R12.Intl_1 := "AlwaysTRUE" AND (("Valves Data".R12_XV02.STATUS = 1) OR ("Valves Data".R12_XV03.STATUS = 1) OR ("Valves Data".R12_XV04.STATUS = 1));
END_REGION

REGION Network 123: R12_XV02
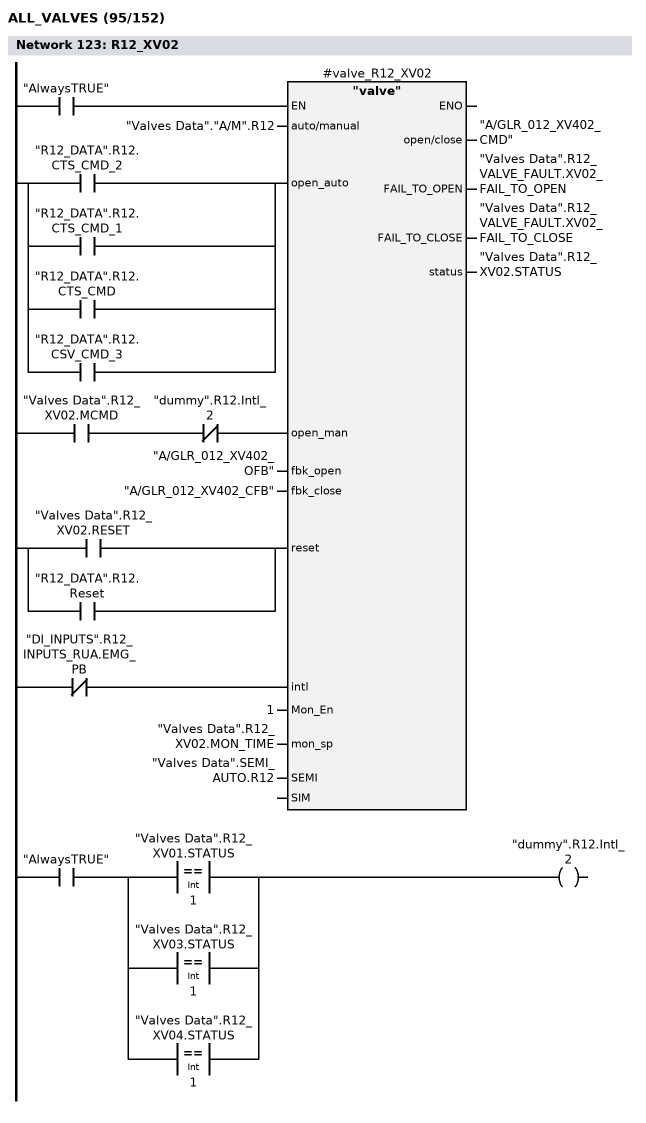
   RUNG wire#powerrail
      Contact( "AlwaysTRUE" )
      #valve_R12_XV02(open_auto := wire#w1, open_man := wire#w2, reset := wire#w3, intl := wire#w4, "auto/manual" := "Valves Data"."A/M".R12, fbk_open := "A/GLR_012_XV402_OFB", fbk_close := "A/GLR_012_XV402_CFB", Mon_En := 1, mon_sp := "Valves Data".R12_XV02.MON_TIME, SEMI := "Valves Data".SEMI_AUTO.R12, SIM :=, "open/close" => "A/GLR_012_XV402_CMD", FAIL_TO_OPEN => "Valves Data".R12_VALVE_FAULT.XV02_FAIL_TO_OPEN, FAIL_TO_CLOSE => "Valves Data".R12_VALVE_FAULT.XV02_FAIL_TO_CLOSE, status => "Valves Data".R12_XV02.STATUS)
   END_RUNG
   RUNG wire#powerrail
      Contact( "R12_DATA".R12.CTS_CMD_2 )
   END_RUNG wire#w1
   RUNG wire#powerrail
      Contact( "R12_DATA".R12.CTS_CMD_1 )
   END_RUNG wire#w1
   RUNG wire#powerrail
      Contact( "R12_DATA".R12.CTS_CMD )
   END_RUNG wire#w1
   RUNG wire#powerrail
      Contact( "R12_DATA".R12.CSV_CMD_3 )
   END_RUNG wire#w1
   RUNG wire#powerrail
      Contact( "Valves Data".R12_XV02.MCMD )
      I_Contact( "dummy".R12.Intl_2 )
   END_RUNG wire#w2
   RUNG wire#powerrail
      Contact( "Valves Data".R12_XV02.RESET )
   END_RUNG wire#w3
   RUNG wire#powerrail
      Contact( "R12_DATA".R12.Reset )
   END_RUNG wire#w3
   RUNG wire#powerrail
      I_Contact( "DI_INPUTS".R12_INPUTS_RUA.EMG_PB )
   END_RUNG wire#w4
   RUNG wire#powerrail
      Contact( "AlwaysTRUE" )
      wire#w5
      { S7_Templates := "SrcType := Int" } EQ_Contact(in1 := "Valves Data".R12_XV01.STATUS, in2 := 1)
      wire#w6
      Coil( "dummy".R12.Intl_2 )
   END_RUNG
   RUNG wire#w5
      { S7_Templates := "SrcType := Int" } EQ_Contact(in1 := "Valves Data".R12_XV03.STATUS, in2 := 1)
   END_RUNG wire#w6
   RUNG wire#w5
      { S7_Templates := "SrcType := Int" } EQ_Contact(in1 := "Valves Data".R12_XV04.STATUS, in2 := 1)
   END_RUNG wire#w6
   // the same network as SCL:
   IF "AlwaysTRUE" THEN
       #valve_R12_XV02("auto/manual" := "Valves Data"."A/M".R12,   // "valve"
                       open_auto := "R12_DATA".R12.CTS_CMD_2 OR "R12_DATA".R12.CTS_CMD_1 OR "R12_DATA".R12.CTS_CMD OR "R12_DATA".R12.CSV_CMD_3,
                       open_man := "Valves Data".R12_XV02.MCMD AND NOT "dummy".R12.Intl_2,
                       fbk_open := "A/GLR_012_XV402_OFB",
                       fbk_close := "A/GLR_012_XV402_CFB",
                       reset := "Valves Data".R12_XV02.RESET OR "R12_DATA".R12.Reset,
                       intl := NOT "DI_INPUTS".R12_INPUTS_RUA.EMG_PB,
                       Mon_En := 1,
                       mon_sp := "Valves Data".R12_XV02.MON_TIME,
                       SEMI := "Valves Data".SEMI_AUTO.R12,
                       "open/close" => "A/GLR_012_XV402_CMD",
                       FAIL_TO_OPEN => "Valves Data".R12_VALVE_FAULT.XV02_FAIL_TO_OPEN,
                       FAIL_TO_CLOSE => "Valves Data".R12_VALVE_FAULT.XV02_FAIL_TO_CLOSE,
                       status => "Valves Data".R12_XV02.STATUS);
   END_IF;
   "dummy".R12.Intl_2 := "AlwaysTRUE" AND (("Valves Data".R12_XV01.STATUS = 1) OR ("Valves Data".R12_XV03.STATUS = 1) OR ("Valves Data".R12_XV04.STATUS = 1));
END_REGION

REGION Network 124: R12_XV03
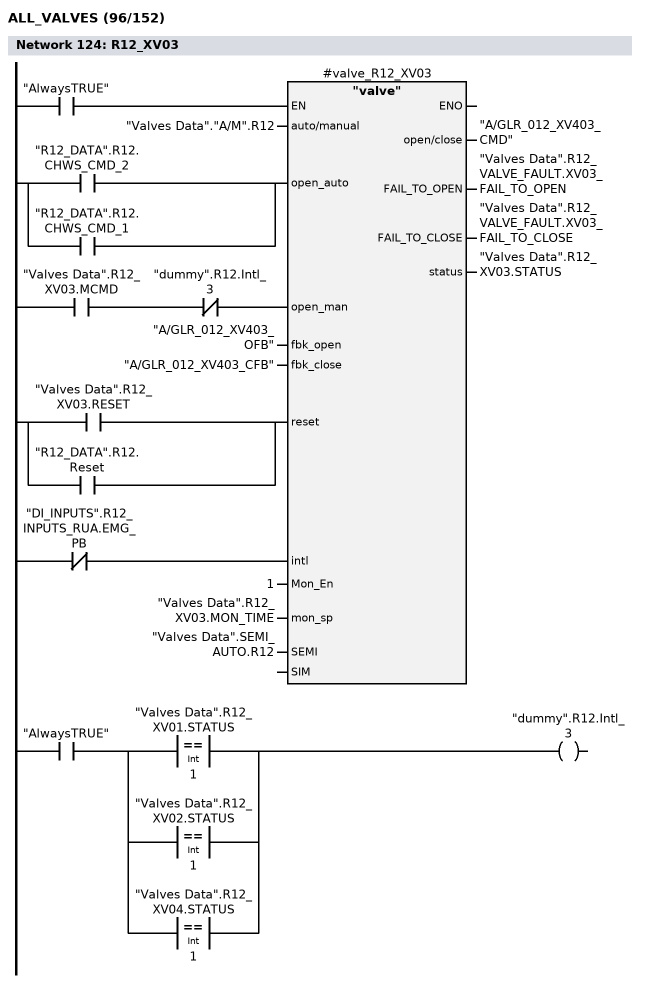
   RUNG wire#powerrail
      Contact( "AlwaysTRUE" )
      #valve_R12_XV03(open_auto := wire#w1, open_man := wire#w2, reset := wire#w3, intl := wire#w4, "auto/manual" := "Valves Data"."A/M".R12, fbk_open := "A/GLR_012_XV403_OFB", fbk_close := "A/GLR_012_XV403_CFB", Mon_En := 1, mon_sp := "Valves Data".R12_XV03.MON_TIME, SEMI := "Valves Data".SEMI_AUTO.R12, SIM :=, "open/close" => "A/GLR_012_XV403_CMD", FAIL_TO_OPEN => "Valves Data".R12_VALVE_FAULT.XV03_FAIL_TO_OPEN, FAIL_TO_CLOSE => "Valves Data".R12_VALVE_FAULT.XV03_FAIL_TO_CLOSE, status => "Valves Data".R12_XV03.STATUS)
   END_RUNG
   RUNG wire#powerrail
      Contact( "R12_DATA".R12.CHWS_CMD_2 )
   END_RUNG wire#w1
   RUNG wire#powerrail
      Contact( "R12_DATA".R12.CHWS_CMD_1 )
   END_RUNG wire#w1
   RUNG wire#powerrail
      Contact( "Valves Data".R12_XV03.MCMD )
      I_Contact( "dummy".R12.Intl_3 )
   END_RUNG wire#w2
   RUNG wire#powerrail
      Contact( "Valves Data".R12_XV03.RESET )
   END_RUNG wire#w3
   RUNG wire#powerrail
      Contact( "R12_DATA".R12.Reset )
   END_RUNG wire#w3
   RUNG wire#powerrail
      I_Contact( "DI_INPUTS".R12_INPUTS_RUA.EMG_PB )
   END_RUNG wire#w4
   RUNG wire#powerrail
      Contact( "AlwaysTRUE" )
      wire#w5
      { S7_Templates := "SrcType := Int" } EQ_Contact(in1 := "Valves Data".R12_XV01.STATUS, in2 := 1)
      wire#w6
      Coil( "dummy".R12.Intl_3 )
   END_RUNG
   RUNG wire#w5
      { S7_Templates := "SrcType := Int" } EQ_Contact(in1 := "Valves Data".R12_XV02.STATUS, in2 := 1)
   END_RUNG wire#w6
   RUNG wire#w5
      { S7_Templates := "SrcType := Int" } EQ_Contact(in1 := "Valves Data".R12_XV04.STATUS, in2 := 1)
   END_RUNG wire#w6
   // the same network as SCL:
   IF "AlwaysTRUE" THEN
       #valve_R12_XV03("auto/manual" := "Valves Data"."A/M".R12,   // "valve"
                       open_auto := "R12_DATA".R12.CHWS_CMD_2 OR "R12_DATA".R12.CHWS_CMD_1,
                       open_man := "Valves Data".R12_XV03.MCMD AND NOT "dummy".R12.Intl_3,
                       fbk_open := "A/GLR_012_XV403_OFB",
                       fbk_close := "A/GLR_012_XV403_CFB",
                       reset := "Valves Data".R12_XV03.RESET OR "R12_DATA".R12.Reset,
                       intl := NOT "DI_INPUTS".R12_INPUTS_RUA.EMG_PB,
                       Mon_En := 1,
                       mon_sp := "Valves Data".R12_XV03.MON_TIME,
                       SEMI := "Valves Data".SEMI_AUTO.R12,
                       "open/close" => "A/GLR_012_XV403_CMD",
                       FAIL_TO_OPEN => "Valves Data".R12_VALVE_FAULT.XV03_FAIL_TO_OPEN,
                       FAIL_TO_CLOSE => "Valves Data".R12_VALVE_FAULT.XV03_FAIL_TO_CLOSE,
                       status => "Valves Data".R12_XV03.STATUS);
   END_IF;
   "dummy".R12.Intl_3 := "AlwaysTRUE" AND (("Valves Data".R12_XV01.STATUS = 1) OR ("Valves Data".R12_XV02.STATUS = 1) OR ("Valves Data".R12_XV04.STATUS = 1));
END_REGION

REGION Network 125: R12_XV04
